   "PopUps_DB_1".Absolute_Encoder[#HMI_No].AE_Position_1 := "Control_DB".VTD_Sys[#Sys_No].Inputs.AE_Position_1;
   "PopUps_DB_1".Absolute_Encoder[#HMI_No].AE_Position_2 := "Control_DB".VTD_Sys[#Sys_No].Inputs.AE_Position_2;
   "PopUps_DB_1".Absolute_Encoder[#HMI_No].AE_Speed := "Control_DB".VTD_Sys[#Sys_No].Inputs.AE_Speed;
   "PopUps_DB_1".Absolute_Encoder[#HMI_No].AE_Status_1 := "Control_DB".VTD_Sys[#Sys_No].Inputs.AE_Status_1;
   "PopUps_DB_1".Absolute_Encoder[#HMI_No].AE_Status_2 := "Control_DB".VTD_Sys[#Sys_No].Inputs.AE_Status_2;

   //Instruction
   IF NOT "VTD_HMI".Charge_VTD_Commands[#HMI_No] THEN
       "Control_DB".VTD_Sys[#Sys_No].Instruction.Reset := "VTD_HMI".Reset[#HMI_No] OR "Screen_DB_1".Reset_All[#HMI_No];
       "Control_DB".VTD_Sys[#Sys_No].Instruction.Enable := "VTD_HMI".Enable[#HMI_No];
       IF "VTD_HMI".Stop[#HMI_No] THEN
           "Control_DB".VTD_Sys[#Sys_No].Instruction.Stop := TRUE;
       ELSIF "Screen_DB_1".Reset_All[1] OR "VTD_HMI".Reset[#HMI_No] THEN
           "Control_DB".VTD_Sys[#Sys_No].Instruction.Stop := "VTD_HMI".Stop[#HMI_No] := FALSE;
       END_IF;

       IF "Control_DB".VTD_Sys[#Sys_No].Mode <> 3 THEN
           "Control_DB".VTD_Sys[#Sys_No].Instruction.Pallet_Type := "VTD_HMI".Pallet_Type[#HMI_No];
           "Control_DB".VTD_Sys[#Sys_No].Instruction.Task_ID := "VTD_HMI".Task_ID[#HMI_No];

           IF "Control_DB".VTD_Sys[#Sys_No].Mode = 2 AND "VTD_HMI".Move_To_Level[#HMI_No] <> 0 THEN
               "Control_DB".VTD_Sys[#Sys_No].Instruction.Move_To_Level := "VTD_HMI".Move_To_Level[#HMI_No];
               "VTD_HMI".Move_To_Level[#HMI_No] := 0;
           END_IF;

           //UP
           IF "Control_DB".VTD_Sys[#Sys_No].LE < "Settings_DB".VTD_Sys[#Sys_No].Teach_Values.Levels_LE[#HMI_Box MOD 10 + 1] - 150
           THEN
               "Control_DB".VTD_Sys[#Sys_No].Instruction.Manual_Up := "VTD_HMI".Manual_Up[#HMI_No];
           ELSE
               "Control_DB".VTD_Sys[#Sys_No].Instruction.Manual_Up := "VTD_HMI".Manual_Up[#HMI_No] := FALSE;
           END_IF;
           //DOWN
           IF "Control_DB".VTD_Sys[#Sys_No].LE > "Settings_DB".VTD_Sys[#Sys_No].Teach_Values.Levels_LE[#HMI_Box MOD 10]
           THEN
               "Control_DB".VTD_Sys[#Sys_No].Instruction.Manual_Down := "VTD_HMI".Manual_Down[#HMI_No];
           ELSE
               "Control_DB".VTD_Sys[#Sys_No].Instruction.Manual_Down := "VTD_HMI".Manual_Down[#HMI_No] := FALSE;
           END_IF;

           "Control_DB".VTD_Sys[#Sys_No].Instruction.Manual_LP_Retract := "VTD_HMI".Manual_DP_Retract[#HMI_No];
           "Control_DB".VTD_Sys[#Sys_No].Instruction.Manual_LP_Extend := "VTD_HMI".Manual_DP_Extend[#HMI_No];
       END_IF;

       //ABSOLUTE ENCODER
       "Control_DB".VTD_Sys[#Sys_No].Outputs.AE_Control_Word_1 := "PopUps_DB_1".Absolute_Encoder[#HMI_No].AE_Control_Word_1;
       "Control_DB".VTD_Sys[#Sys_No].Outputs.AE_Control_Word_2 := "PopUps_DB_1".Absolute_Encoder[#HMI_No].AE_Control_Word_2;

       //LINEAR ENCODER
       "VTD_HMI".LE_Bypass[#Sys_No] := "PopUps_DB_1".Linear_Encoder[#HMI_No].LE_Bypass;

       //BARCODE
       #BCD_Start_Comm_Test_HMI := "PopUps_DB_1".Lector_Barcode[#HMI_No].BCD_Test_Comm;
       #BCD_Enable_Trigger_HMI  := "PopUps_DB_1".Lector_Barcode[#HMI_No].BCD_Enable_Trigger;
       #BCD_Disable_Trigger_HMI   := "PopUps_DB_1".Lector_Barcode[#HMI_No].BCD_Disable_Trigger;
       #BCD_Execute_Function  := "PopUps_DB_1".Lector_Barcode[#HMI_No].BCD_Execute_Function;
   END_IF;
END_FUNCTION

FUNCTION "FindBoolField" : Bool   // FC17, SCL
{ S7_Optimized_Access := 'TRUE' }
VERSION : 0.1
// stored: AutoNumber true, IsIECCheckEnabled false, SetENOAutomatically false, UDAEnableTagReadback false
   VAR_INPUT
      FieldName : String;
      JsonStr : String;
   END_VAR
   VAR_TEMP
      searchStr : String;
      foundPos : Int;
      valueStr : String;
      afterField : String;
      bResult : Bool;
   END_VAR
BEGIN
   // Build search string
   #searchStr := CONCAT(IN1 := '"', IN2 := #FieldName);
   #searchStr := CONCAT(IN1 := #searchStr, IN2 := '" :');

   // Serach for JSON field
   #foundPos := FIND(IN1 := #JsonStr, IN2 := #searchStr);

   IF #foundPos > 0 THEN
       // Take to 20 characters after the field
       #afterField := MID(IN := #JsonStr, P := #foundPos + LEN(#searchStr), L := 20);

       // Normalize to remove whitespace if necessary
       // (or compare directly)
       IF FIND(IN1 := #afterField, IN2 := 'true') > 0 THEN
           #bResult := TRUE;
       ELSIF FIND(IN1 := #afterField, IN2 := 'false') > 0 THEN
           #bResult := FALSE;
       ELSE
           #bResult := FALSE; // default if value not found
       END_IF;
   ELSE
       #bResult := FALSE;
   END_IF;

   #FindBoolField := #bResult;
END_FUNCTION

FUNCTION "FindDINTFieldFragmented" : DInt   // FC20, SCL
{ S7_Optimized_Access := 'TRUE' }
VERSION : 0.1
// stored: AutoNumber true, IsIECCheckEnabled false, SetENOAutomatically false, UDAEnableTagReadback false
   VAR_INPUT
      FieldName : String;
      Str1 : String;
      Str2 : String;
   END_VAR
   VAR_TEMP
      searchStr : String;
      iStart : Int;
      iEnd : Int;
      tempVal : String;
      fieldFound : Bool;
      loopIdx : Int;
   END_VAR
BEGIN
   // Build search string
   #searchStr := CONCAT(IN1 := '"', IN2 := #FieldName);
   #searchStr := CONCAT(IN1 := #searchStr, IN2 := '" :');

   // Serach for JSON field
   #iStart := FIND(IN1 := #Str1, IN2 := #searchStr);

   IF #iStart > 0 THEN
       // Found full field in String_1
       #iEnd := FIND(IN1 := MID(IN := #Str1, P := #iStart + LEN(#searchStr), L := 20), IN2 := ',');
       IF #iEnd = 0 THEN
           #iEnd := FIND(IN1 := MID(IN := #Str1, P := #iStart + LEN(#searchStr), L := 20), IN2 := '}');
       END_IF;
       IF #iEnd > 0 THEN
           #tempVal := MID(IN := #Str1, P := #iStart + LEN(#searchStr), L := #iEnd - 1);
           #fieldFound := TRUE;
       END_IF;
   END_IF;

   // Search for full field in Str2
   IF NOT #fieldFound THEN
       #iStart := FIND(IN1 := #Str2, IN2 := #searchStr);
       IF #iStart > 0 THEN
           #iEnd := FIND(IN1 := MID(IN := #Str2, P := #iStart + LEN(#searchStr), L := 20), IN2 := ',');
           IF #iEnd = 0 THEN
               #iEnd := FIND(IN1 := MID(IN := #Str2, P := #iStart + LEN(#searchStr), L := 20), IN2 := '}');
           END_IF;
           IF #iEnd > 0 THEN
               #tempVal := MID(IN := #Str2, P := #iStart + LEN(#searchStr), L := #iEnd - 1);
               #fieldFound := TRUE;
           END_IF;
       END_IF;
   END_IF;

   // Search for fragmented field: end of name in Str1 and beginning in Str2
   IF NOT #fieldFound THEN
       // Examines last 10 characters of String_1
       FOR #loopIdx := LEN(#Str1) - 15 TO LEN(#Str1) DO
           IF MID(IN := #Str1, P := #loopIdx, L := 1) = '"' THEN
               #tempVal := MID(IN := #Str1, P := #loopIdx, L := LEN(#Str1) - #loopIdx + 1);
               #tempVal := CONCAT(IN1 := #tempVal, IN2 := #Str2); // concatenates piece from beginning of String_2
               #iStart := FIND(IN1 := #tempVal, IN2 := #searchStr);
               IF #iStart > 0 THEN
                   #iEnd := FIND(IN1 := MID(IN := #tempVal, P := #iStart + LEN(#searchStr), L := 20), IN2 := ',');
                   IF #iEnd = 0 THEN
                       #iEnd := FIND(IN1 := MID(IN := #tempVal, P := #iStart + LEN(#searchStr), L := 20), IN2 := '}');
                   END_IF;
                   IF #iEnd > 0 THEN
                       #tempVal := MID(IN := #tempVal, P := #iStart + LEN(#searchStr), L := #iEnd - 1);
                       #fieldFound := TRUE;
                   END_IF;
               END_IF;
               EXIT; // found, you can leave
           END_IF;
       END_FOR;
   END_IF;

   // Return value
   IF #fieldFound THEN
       #FindDINTFieldFragmented := STRING_TO_DINT(#tempVal);
   ELSE
       #FindDINTFieldFragmented := -9999; // default value if not found
   END_IF;
END_FUNCTION

FUNCTION "FindINTFieldFragmented" : Int   // FC22, SCL
{ S7_Optimized_Access := 'TRUE' }
VERSION : 0.1
// stored: AutoNumber true, IsIECCheckEnabled false, SetENOAutomatically false, UDAEnableTagReadback false
   VAR_INPUT
      FieldName : String;
      Str1 : String;
      Str2 : String;
   END_VAR
   VAR_TEMP
      searchStr : String;
      iStart : Int;
      iEnd : Int;
      tempVal : String;
      fieldFound : Bool;
      loopIdx : Int;
   END_VAR
BEGIN
   // Build search string
   #searchStr := CONCAT(IN1 := '"', IN2 := #FieldName);
   #searchStr := CONCAT(IN1 := #searchStr, IN2 := '" :');

   // Serach for JSON field
   #iStart := FIND(IN1 := #Str1, IN2 := #searchStr);

   IF #iStart > 0 THEN
       // Found full field in String_1
       #iEnd := FIND(IN1 := MID(IN := #Str1, P := #iStart + LEN(#searchStr), L := 20), IN2 := ',');
       IF #iEnd = 0 THEN
           #iEnd := FIND(IN1 := MID(IN := #Str1, P := #iStart + LEN(#searchStr), L := 20), IN2 := '}');
       END_IF;
       IF #iEnd > 0 THEN
           #tempVal := MID(IN := #Str1, P := #iStart + LEN(#searchStr), L := #iEnd - 1);
           #fieldFound := TRUE;
       END_IF;
   END_IF;

   // Search for full field in Str2
   IF NOT #fieldFound THEN
       #iStart := FIND(IN1 := #Str2, IN2 := #searchStr);
       IF #iStart > 0 THEN
           #iEnd := FIND(IN1 := MID(IN := #Str2, P := #iStart + LEN(#searchStr), L := 20), IN2 := ',');
           IF #iEnd = 0 THEN
               #iEnd := FIND(IN1 := MID(IN := #Str2, P := #iStart + LEN(#searchStr), L := 20), IN2 := '}');
           END_IF;
           IF #iEnd > 0 THEN
               #tempVal := MID(IN := #Str2, P := #iStart + LEN(#searchStr), L := #iEnd - 1);
               #fieldFound := TRUE;
           END_IF;
       END_IF;
   END_IF;

   // Search for fragmented field: end of name in Str1 and beginning in Str2
   IF NOT #fieldFound THEN
       // Examines last 10 characters of String_1
       FOR #loopIdx := LEN(#Str1) - 15 TO LEN(#Str1) DO
           IF MID(IN := #Str1, P := #loopIdx, L := 1) = '"' THEN
               #tempVal := MID(IN := #Str1, P := #loopIdx, L := LEN(#Str1) - #loopIdx + 1);
               #tempVal := CONCAT(IN1 := #tempVal, IN2 := #Str2); // concatenates piece from beginning of String_2
               #iStart := FIND(IN1 := #tempVal, IN2 := #searchStr);
               IF #iStart > 0 THEN
                   #iEnd := FIND(IN1 := MID(IN := #tempVal, P := #iStart + LEN(#searchStr), L := 20), IN2 := ',');
                   IF #iEnd = 0 THEN
                       #iEnd := FIND(IN1 := MID(IN := #tempVal, P := #iStart + LEN(#searchStr), L := 20), IN2 := '}');
                   END_IF;
                   IF #iEnd > 0 THEN
                       #tempVal := MID(IN := #tempVal, P := #iStart + LEN(#searchStr), L := #iEnd - 1);
                       #fieldFound := TRUE;
                   END_IF;
               END_IF;
               EXIT; // found, you can leave
           END_IF;
       END_FOR;
   END_IF;

   // Return value
   IF #fieldFound THEN
       #FindINTFieldFragmented := STRING_TO_INT(#tempVal);
   ELSE
       #FindINTFieldFragmented := -9999; // default value if not found
   END_IF;
END_FUNCTION

FUNCTION "FindIntField" : Int   // FC18, SCL
{ S7_Optimized_Access := 'TRUE' }
VERSION : 0.1
// stored: AutoNumber true, IsIECCheckEnabled false, SetENOAutomatically false, UDAEnableTagReadback false
   VAR_INPUT
      FieldName : String;
      JsonStr : String;
   END_VAR
   VAR_TEMP
      searchStr : String;
      foundPos : Int;
      valueStr : String;
      delimPos : Int;
   END_VAR
BEGIN
   // Set up the search pattern, e.g. '"id":'
   #searchStr := CONCAT(IN1 := '"', IN2 := #FieldName);
   #searchStr := CONCAT(IN1 := #searchStr, IN2 := '" :');

   // Search the field
   #foundPos := FIND(IN1 := #JsonStr, IN2 := #searchStr);

   IF #foundPos > 0 THEN
       // Try to find a comma after the value
       #delimPos := FIND(
                         IN1 := MID(IN := #JsonStr, P := #foundPos + LEN(#searchStr), L := 10),
                         IN2 := ','
       );

       // If there is no comma, try to find the closing brace '}'
       IF #delimPos = 0 THEN
           #delimPos := FIND(
                             IN1 := MID(IN := #JsonStr, P := #foundPos + LEN(#searchStr), L := 10),
                             IN2 := '}'
           );
       END_IF;

       // If you find the end of value, extract the value
       IF #delimPos > 0 THEN
           #valueStr := MID(
                            IN := #JsonStr,
                            P := #foundPos + LEN(#searchStr),
                            L := #delimPos - 1
           );
           #FindIntField := STRING_TO_INT(#valueStr);
           RETURN;
       END_IF;
   END_IF;

   // Default return if not found or error
   #FindIntField := -9999;
END_FUNCTION

FUNCTION "FindSTRINGFieldFragmented" : String   // FC21, SCL
{ S7_Optimized_Access := 'TRUE' }
VERSION : 0.1
// stored: AutoNumber true, IsIECCheckEnabled false, SetENOAutomatically false, UDAEnableTagReadback false
   VAR_INPUT
      FieldName : String;
      Str1 : String;
      Str2 : String;
   END_VAR
   VAR_TEMP
      searchStr : String;
      iStart : Int;
      iEnd : Int;
      tempVal : String;
      fieldFound : Bool;
      loopIdx : Int;
   END_VAR
BEGIN
   // Build search string
   #searchStr := CONCAT(IN1 := '"', IN2 := #FieldName);
   #searchStr := CONCAT(IN1 := #searchStr, IN2 := '" :');

   // Serach for JSON field
   #iStart := FIND(IN1 := #Str1, IN2 := #searchStr);

   IF #iStart > 0 THEN
       // Found full field in String_1
       #iEnd := FIND(IN1 := MID(IN := #Str1, P := #iStart + LEN(#searchStr), L := 20), IN2 := ',');
       IF #iEnd = 0 THEN
           #iEnd := FIND(IN1 := MID(IN := #Str1, P := #iStart + LEN(#searchStr), L := 20), IN2 := '}');
       END_IF;
       IF #iEnd > 0 THEN
           #tempVal := MID(IN := #Str1, P := #iStart + LEN(#searchStr), L := #iEnd - 1);
           #fieldFound := TRUE;
       END_IF;
   END_IF;

   // Search for full field in Str2
   IF NOT #fieldFound THEN
       #iStart := FIND(IN1 := #Str2, IN2 := #searchStr);
       IF #iStart > 0 THEN
           #iEnd := FIND(IN1 := MID(IN := #Str2, P := #iStart + LEN(#searchStr), L := 20), IN2 := ',');
           IF #iEnd = 0 THEN
               #iEnd := FIND(IN1 := MID(IN := #Str2, P := #iStart + LEN(#searchStr), L := 20), IN2 := '}');
           END_IF;
           IF #iEnd > 0 THEN
               #tempVal := MID(IN := #Str2, P := #iStart + LEN(#searchStr), L := #iEnd - 1);
               #fieldFound := TRUE;
           END_IF;
       END_IF;
   END_IF;

   // Search for fragmented field: end of name in Str1 and beginning in Str2
   IF NOT #fieldFound THEN
       // Examines last 10 characters of String_1
       FOR #loopIdx := LEN(#Str1) - 15 TO LEN(#Str1) DO
           IF MID(IN := #Str1, P := #loopIdx, L := 1) = '"' THEN
               #tempVal := MID(IN := #Str1, P := #loopIdx, L := LEN(#Str1) - #loopIdx + 1);
               #tempVal := CONCAT(IN1 := #tempVal, IN2 := #Str2); // concatenates piece from beginning of String_2
               #iStart := FIND(IN1 := #tempVal, IN2 := #searchStr);
               IF #iStart > 0 THEN
                   #iEnd := FIND(IN1 := MID(IN := #tempVal, P := #iStart + LEN(#searchStr), L := 20), IN2 := ',');
                   IF #iEnd = 0 THEN
                       #iEnd := FIND(IN1 := MID(IN := #tempVal, P := #iStart + LEN(#searchStr), L := 20), IN2 := '}');
                   END_IF;
                   IF #iEnd > 0 THEN
                       #tempVal := MID(IN := #tempVal, P := #iStart + LEN(#searchStr), L := #iEnd - 1);
                       #fieldFound := TRUE;
                   END_IF;
               END_IF;
               EXIT; // found, you can leave
           END_IF;
       END_FOR;
   END_IF;

   // Return value
   IF #fieldFound THEN
       #FindSTRINGFieldFragmented := #tempVal;
   ELSE
       #FindSTRINGFieldFragmented := 'NOT FOUND'; // default value if not found
   END_IF;
END_FUNCTION

FUNCTION "FindStringField" : String   // FC19, SCL
{ S7_Optimized_Access := 'TRUE' }
VERSION : 0.1
// stored: AutoNumber true, IsIECCheckEnabled false, SetENOAutomatically false, UDAEnableTagReadback false
   VAR_INPUT
      FieldName : String;
      JsonStr : String;
   END_VAR
   VAR_TEMP
      searchStr : String;
      foundPos : Int;
      resultStr : String;
      quotePos1 : Int;
      quotePos2 : Int;
   END_VAR
BEGIN
   // Sets search pattern → ex: '"loadstate":'
   #searchStr := CONCAT(IN1 := '"', IN2 := #FieldName);
   #searchStr := CONCAT(IN1 := #searchStr, IN2 := '" :');

   // Search in JSON
   #foundPos := FIND(IN1 := #JsonStr, IN2 := #searchStr);

   IF #foundPos > 0 THEN
       // Finds first quote after field
       #quotePos1 := FIND(IN1 := MID(IN := #JsonStr, P := #foundPos + LEN(#searchStr), L := 20), IN2 := '"');

       IF #quotePos1 > 0 THEN
           // Finds second quote after the first
           #quotePos2 := FIND(
                              IN1 := MID(IN := #JsonStr, P := #foundPos + LEN(IN := #searchStr) + #quotePos1, L := 10),
                              IN2 := '"'
           );

           IF #quotePos2 > 0 THEN
               #resultStr := MID(
                                 IN := #JsonStr,
                                 P := #foundPos + LEN(#searchStr) + #quotePos1,
                                 L := #quotePos2 - 1
               );
               #FindStringField := #resultStr;
               RETURN;
           END_IF;
       END_IF;
   END_IF;

   // If not found, returns empty string
   #FindStringField := '';
END_FUNCTION

FUNCTION "Gate_Status_Update_FC" : Void   // FC49, SCL
{ S7_Optimized_Access := 'TRUE' }
VERSION : 0.1
// stored: AutoNumber true, IsIECCheckEnabled false, SetENOAutomatically false, UDAEnableTagReadback false
   VAR_INPUT
      Gate_Index : Int;
      Request_Access : Bool;
      Stop_Mode_Granted : Bool;
   END_VAR
   VAR_OUTPUT
      DB_SM_To_LGX_Gate_Status : Array[0..10] of Byte;
   END_VAR
   VAR_TEMP
      tGateByte : Byte;
   END_VAR
BEGIN
   #tGateByte := 0;

   IF #Request_Access THEN
       #tGateByte := #tGateByte OR BYTE#16#01;
   END_IF; // Bit 0
   IF #Stop_Mode_Granted THEN
       #tGateByte := #tGateByte OR BYTE#16#02;
   END_IF; // Bit 1
   // Bits 2..7: Free

   IF #Gate_Index >= 0 AND #Gate_Index <= 10 THEN
       #DB_SM_To_LGX_Gate_Status[#Gate_Index] := #tGateByte;
   END_IF;
END_FUNCTION

FUNCTION "HMI_SAFETY_FC" : Void   // FC43, F_FBD
{ S7_Optimized_Access := 'TRUE' }
VERSION : 0.1
// stored: AutoNumber true, IsIECCheckEnabled false, UDAEnableTagReadback false
   VAR_INPUT
      HMI_Box_Connected : Int;
      HMI_Reset : Bool;
      HMI_EStop : Bool;
      HMI_Profinet_Error : Bool;
      Local_Mode : Bool;
   END_VAR
   VAR_OUTPUT
      HMI_Estop_Pressed_1 : Bool;
      HMI_Estop_Pressed_2 : Bool;
      HMI_Estop_Pressed_3 : Bool;
      HMI_Estop_Pressed_4 : Bool;
      HMI_Estop_Pressed_5 : Bool;
      Reset_Comissioning_1 : Bool;
      Reset_Comissioning_2 : Bool;
      Reset_Comissioning_3 : Bool;
      Reset_Comissioning_4 : Bool;
      Reset_Comissioning_5 : Bool;
   END_VAR
   VAR_TEMP   // added for the SCL form of the ladder/FBD networks
      _w1 : Bool;
   END_VAR
BEGIN

REGION Network 1: HMI CONNECTED IN THE SYSTEM 1
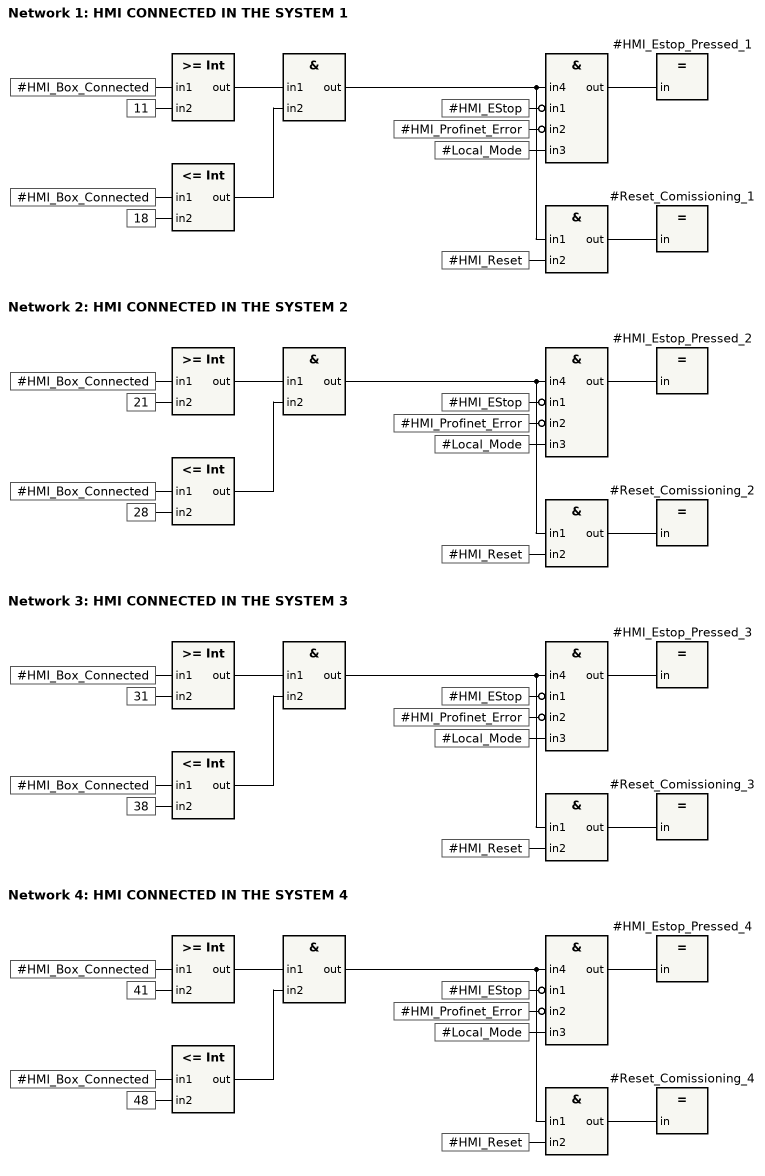
   #_w1 := (#HMI_Box_Connected >= 11) AND (#HMI_Box_Connected <= 18);
   #HMI_Estop_Pressed_1 := #_w1 AND NOT #HMI_EStop AND NOT #HMI_Profinet_Error AND #Local_Mode;
   #Reset_Comissioning_1 := #_w1 AND #HMI_Reset;
END_REGION

REGION Network 2: HMI CONNECTED IN THE SYSTEM 2
   #_w1 := (#HMI_Box_Connected >= 21) AND (#HMI_Box_Connected <= 28);
   #HMI_Estop_Pressed_2 := #_w1 AND NOT #HMI_EStop AND NOT #HMI_Profinet_Error AND #Local_Mode;
   #Reset_Comissioning_2 := #_w1 AND #HMI_Reset;
END_REGION

REGION Network 3: HMI CONNECTED IN THE SYSTEM 3
   #_w1 := (#HMI_Box_Connected >= 31) AND (#HMI_Box_Connected <= 38);
   #HMI_Estop_Pressed_3 := #_w1 AND NOT #HMI_EStop AND NOT #HMI_Profinet_Error AND #Local_Mode;
   #Reset_Comissioning_3 := #_w1 AND #HMI_Reset;
END_REGION

REGION Network 4: HMI CONNECTED IN THE SYSTEM 4
   #_w1 := (#HMI_Box_Connected >= 41) AND (#HMI_Box_Connected <= 48);
   #HMI_Estop_Pressed_4 := #_w1 AND NOT #HMI_EStop AND NOT #HMI_Profinet_Error AND #Local_Mode;
   #Reset_Comissioning_4 := #_w1 AND #HMI_Reset;
END_REGION

REGION Network 5: HMI CONNECTED IN THE SYSTEM 5
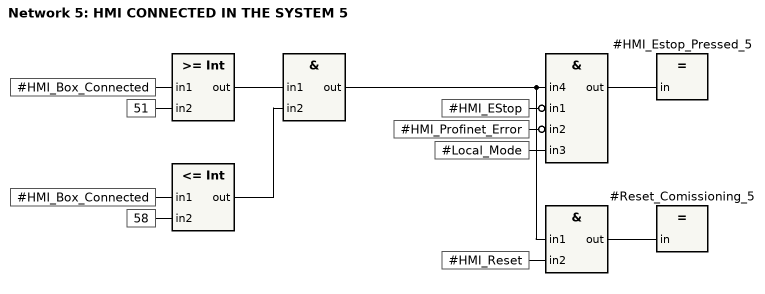
   #_w1 := (#HMI_Box_Connected >= 51) AND (#HMI_Box_Connected <= 58);
   #HMI_Estop_Pressed_5 := #_w1 AND NOT #HMI_EStop AND NOT #HMI_Profinet_Error AND #Local_Mode;
   #Reset_Comissioning_5 := #_w1 AND #HMI_Reset;
END_REGION
END_FUNCTION

FUNCTION "Handshake_Infeed_FC" : Void   // FC47, SCL
{ S7_Optimized_Access := 'TRUE' }
VERSION : 0.1
// stored: AutoNumber true, IsIECCheckEnabled false, SetENOAutomatically false, UDAEnableTagReadback false
   VAR_INPUT
      Infeed_Stop_Sensor : Bool;
      Ready_To_Receive : Bool;
      Auto_Mode : Bool;
      Transfer_In_Progress : Bool;
      DB_LGX_To_SM_Infeed_Ready_To_Send : Bool;
      DB_LGX_To_SM_Infeed_Transfer_In_Progress : Bool;
   END_VAR
   VAR_OUTPUT
      Fault_Handshake : Bool;
      DB_SM_To_LGX_Infeed_Ready_To_Receive : Bool;
      DB_SM_To_LGX_Infeed_Pallet_Received : Bool;
      DB_SM_To_LGX_Infeed_Transfer_In_Progress : Bool;
   END_VAR
   VAR_TEMP
      tReady_To_Receive_Condition : Bool;
      tPallet_Received_Condition : Bool;
   END_VAR
BEGIN
   // ---------------------------------------------------------
   // STEP 1: Is SM ready to receive?
   // Condition: SM in Auto, infeed conveyor healthy,
   //            no transfer in progress, no alarm
   // ---------------------------------------------------------
   #tReady_To_Receive_Condition :=
   #Auto_Mode
   AND #Ready_To_Receive
   AND NOT #DB_SM_To_LGX_Infeed_Ready_To_Receive
   AND NOT #DB_SM_To_LGX_Infeed_Pallet_Received;

   IF #DB_LGX_To_SM_Infeed_Ready_To_Send
       AND #tReady_To_Receive_Condition THEN
       #DB_SM_To_LGX_Infeed_Ready_To_Receive := TRUE;
   END_IF;

   // ---------------------------------------------------------
   // STEP 2: Confirm pallet received
   // Condition: Photocell active while transfer is in progress
   // ---------------------------------------------------------
   // #tPallet_Received_Condition :=
   // #Infeed_Stop_Sensor
   // AND #DB_LGX_To_SM_Infeed_Transfer_In_Progress
   // AND #DB_SM_To_LGX_Infeed_Ready_To_Receive;
   // 
   #tPallet_Received_Condition :=
   #Infeed_Stop_Sensor;

   IF #tPallet_Received_Condition THEN
       #DB_SM_To_LGX_Infeed_Pallet_Received := TRUE;
       #DB_SM_To_LGX_Infeed_Ready_To_Receive := FALSE;
   ELSE
       #DB_SM_To_LGX_Infeed_Pallet_Received := FALSE;
   END_IF;

   // ---------------------------------------------------------
   // STEP 3: Reset after LGX confirms end of transfer
   // (LGX resets Transfer_In_Progress upon receiving Pallet_Received)
   // ---------------------------------------------------------
   // IF #DB_SM_To_LGX_Infeed_Pallet_Received
   //     AND NOT #DB_LGX_To_SM_Infeed_Transfer_In_Progress THEN
   //     #DB_SM_To_LGX_Infeed_Pallet_Received := FALSE;
   // END_IF;

   // ---------------------------------------------------------
   // STEP 4: Reset Ready_To_Receive if LGX withdraws Ready_To_Send
   // (e.g. LGX cancelled the operation before starting transfer)
   // ---------------------------------------------------------
   IF NOT #DB_LGX_To_SM_Infeed_Ready_To_Send
       AND NOT #DB_LGX_To_SM_Infeed_Transfer_In_Progress THEN
       #DB_SM_To_LGX_Infeed_Ready_To_Receive := FALSE;
   END_IF;

   // ---------------------------------------------------------
   // FAULT SUPERVISION
   // If Transfer_In_Progress remains active without pallet arriving:
   // use external timer / timeout bit (implement in OB1)
   // ---------------------------------------------------------
   #Fault_Handshake := FALSE; // Placeholder - implement watchdog

   #DB_SM_To_LGX_Infeed_Transfer_In_Progress := #Transfer_In_Progress;
END_FUNCTION

FUNCTION "Handshake_Outfeed_FC" : Void   // FC51, SCL
{ S7_Optimized_Access := 'TRUE' }
VERSION : 0.1
// stored: AutoNumber true, IsIECCheckEnabled false, SetENOAutomatically false, UDAEnableTagReadback false
   VAR_INPUT
      Auto_Mode : Bool;
      Ready_To_Send : Bool;
      Conv_Occupied : Bool;
      Transfer_In_Progress : Bool;
      DB_LGX_To_SM_Outfeed_Ready_To_Receive : Bool;
   END_VAR
   VAR_OUTPUT
      Fault_Handshake : Bool;
      DB_SM_To_LGX_Outfeed_Transfer_In_Progress : Bool;
      DB_SM_To_LGX_Outfeed_Ocuppied : Bool;
      DB_SM_To_LGX_Outfeed_Ready_To_Send : Bool;
   END_VAR
   VAR_TEMP
      tCanSend : Bool;
   END_VAR
BEGIN
   // ---------------------------------------------------------
   // STEP 1: Is SM ready to send?
   // Condition: pallet waiting at exit, SM in auto,
   //            no transfer in progress
   // ---------------------------------------------------------
   #tCanSend :=
   #Auto_Mode
   AND #Conv_Occupied
   AND #Ready_To_Send
   AND NOT #DB_SM_To_LGX_Outfeed_Transfer_In_Progress;

   IF #tCanSend
       AND NOT #DB_SM_To_LGX_Outfeed_Ready_To_Send THEN
       #DB_SM_To_LGX_Outfeed_Ready_To_Send := TRUE;
   END_IF;

   // ---------------------------------------------------------
   // STEP 2: LGX responded Ready_To_Receive → start transfer
   // ---------------------------------------------------------
   IF NOT #Conv_Occupied THEN
       // #DB_SM_To_LGX_Outfeed_Transfer_In_Progress := TRUE;
       #DB_SM_To_LGX_Outfeed_Ready_To_Send := FALSE;
   END_IF;

   // ---------------------------------------------------------
   // STEP 3: LGX confirmed pallet received
   // → SM resets Transfer_In_Progress
   // ---------------------------------------------------------
   // IF #DB_SM_To_LGX_Outfeed_Transfer_In_Progress
   //     AND #DB_LGX_To_SM_Outfeed_Ready_To_Receive THEN
   //     #DB_SM_To_LGX_Outfeed_Transfer_In_Progress := FALSE;
   // END_IF;

   #DB_SM_To_LGX_Outfeed_Transfer_In_Progress := #Transfer_In_Progress;
   #DB_SM_To_LGX_Outfeed_Ocuppied := #Conv_Occupied;
   // ---------------------------------------------------------
   // STEP 4: Reset Ready_To_Send if pallet removed or SM left auto mode
   // ---------------------------------------------------------
   IF NOT #Ready_To_Send OR NOT #Auto_Mode THEN
       IF NOT #DB_SM_To_LGX_Outfeed_Transfer_In_Progress THEN
           #DB_SM_To_LGX_Outfeed_Ready_To_Send := FALSE;
       END_IF;
   END_IF;

   #Fault_Handshake := FALSE; // Placeholder
END_FUNCTION

FUNCTION "ID_Decode_F" : Void   // FC3, SCL
{ S7_Optimized_Access := 'TRUE' }
VERSION : 0.1
// stored: AutoNumber true, IsIECCheckEnabled false, SetENOAutomatically false, UDAEnableTagReadback false
   VAR_INPUT
      ID : DInt;
   END_VAR
   VAR_IN_OUT
      ID_Decoded : "ID_Decoded";
   END_VAR
   VAR_TEMP
      Temp : UInt;
   END_VAR
BEGIN

   // Extract XX (first two digits)
   #ID_Decoded.Device_Type := #ID / 10000;        // 123456 / 10000 = 12

   // Extract YY (middle two digits)
   #ID_Decoded.Level := (#ID MOD 10000) / 100; // 123456 % 10000 = 3456 → 3456 / 100 = 34

   // Extract ZZ (last two digits)
   #ID_Decoded.VTD := #ID MOD 100;       // 123456 % 100 = 56
END_FUNCTION

FUNCTION "IsIPAddress" : Bool   // FC4, SCL
TITLE = IsIPAddress
{ S7_Optimized_Access := 'TRUE' }
VERSION : 0.1
// Evaluates whether a given String contains a valid IP address
// stored: AutoNumber true, IsIECCheckEnabled true, SetENOAutomatically true, UDAEnableTagReadback false
   VAR_INPUT
      address : String;   // Address to be evaluated
   END_VAR
   VAR_OUTPUT
      ipAddress : IP_V4;   // Parsed IP address if passed address is IP address
   END_VAR
   VAR_TEMP
      tempAddress : String;   // Passed address
      tempOctet : String;   // Current octet
      tempIndex : DInt;   // Index for loop
      tempPos : Int;   // Position of found separator
      tempNum : Int;   // Converted octet
      tempIp : IP_V4;   // Parsed IP address
   END_VAR
   VAR CONSTANT
      MAX_VALUE : USInt := 255;   // Max. valid value of octet
      NUM_OCTETS : DInt := 4;   // Number of octets
      CHAR_ZERO : Char := '0';   // ASCII character '0'
   END_VAR
   // Ret_Val : Return value
BEGIN
   REGION BLOCK INFO HEADER
     //===============================================================================
     // SIEMENS / (c)Copyright 2024
     //-------------------------------------------------------------------------------
     // Title:        IsIPAddress
     // Function:     Evaluates whether a given String contains a valid IP address
     // Library:      --
     // Author:       Siemens Industry Online Support
     // Tested with:  CPU 1515-2 PN V3.1
     // Engineering:  TIA Portal V17
     // Restrictions: --
     // Requirements: S7-1200 with firmware V4.4 or higher
     //               S7-1500 with firmware V2.0 or higher
     //-------------------------------------------------------------------------------
     // Change log table:
     // Version  | Date       | Expert in charge       | Changes applied
     //-------------------------------------------------------------------------------
     // 01.00.00 | 2024-02-12 | Online Support         | First released version
     //===============================================================================
   END_REGION

   #tempAddress := #address;
   #IsIPAddress := FALSE; // Will be overwritten if IP address is detected
   #ipAddress := #tempIp; // Zero output parameter

   FOR #tempIndex := 1 TO #NUM_OCTETS DO
     #tempPos := FIND(IN1 := #tempAddress, IN2 := '.'); // Find separator

     IF (#tempPos > 0 OR #tempIndex = #NUM_OCTETS) // Separator found with exception of last octet
       AND NOT (#tempPos > 0 AND #tempIndex = #NUM_OCTETS) // No separator found in last octet
       AND #tempPos <= 4 // 3  characters or less
     THEN
       IF #tempIndex < #NUM_OCTETS THEN // First three octets
         #tempOctet := LEFT(IN := #tempAddress, L := #tempPos - 1);
       ELSE// Last octet
         #tempOctet := #tempAddress;
       END_IF;

       STRG_VAL(IN := #tempOctet,
                FORMAT := 0,
                P := 1,
                OUT => #tempNum);

       IF #tempNum >= 0 AND #tempNum <= #MAX_VALUE // Within 0 and 255
         AND NOT (#tempNum = 0 AND #tempIndex = 1) // Not 0 in first octet
         AND NOT (#tempNum = 0 AND #tempOctet[1] <> #CHAR_ZERO) // Not 0 because of invalid character
       THEN
         #tempIp.ADDR[#tempIndex] := INT_TO_BYTE(#tempNum);
         #tempAddress := RIGHT(IN := #tempAddress, L := LEN(#tempAddress) - #tempPos); // Remove evaluated octet
       ELSE // Address is not IP address
         EXIT;
       END_IF;
     ELSE // Address is not IP address
       EXIT;
     END_IF;

     IF #tempIndex = #NUM_OCTETS THEN // End of loop reached, address is IP address
       #ipAddress := #tempIp;
       #IsIPAddress := true;
     END_IF;
   END_FOR;
END_FUNCTION

FUNCTION "LMQTT_ConvertToUtf8" : Void   // FC6, SCL
TITLE = LMQTT_ConvertToUtf8
{ S7_Optimized_Access := 'TRUE' }
AUTHOR : SIEMENS
FAMILY : LMQTT
VERSION : 1.0
// Function to convert a WCHAR to a UTF-8 conformant byte sequence
// stored: AutoNumber true, IsIECCheckEnabled true, SetENOAutomatically false, UDAEnableTagReadback false
   VAR_INPUT
      character : WChar;   // Character that shall be converted to UTF-8
   END_VAR
   VAR_OUTPUT
      convertedUtf8 : DWord;   // UTF-8 conformant byte sequence. B0 stores first Byte, B1 second and B2 third Byte. B3 is not used
      bytesUsed : USInt;   // Amount of Bytes converted. Ranges from 1 to 3.
      error : Bool;   // TRUE: An error occurred during the execution of the FC
      status : Word;   // 16#0000 - 16#7FFF: Status of the FC, 16#8000 - 16#FFFF: Error identification
   END_VAR
   VAR_TEMP
      tempStatus : Word;   // temp value for output 'status'
      tempConvertedUtf8 : DWord;   // temp value for output 'convertedUtf8'
      tempBytesUsed : USInt;   // temp value for output 'bytesUsed'
      tempCharacter : WChar;   // temp value for input 'character'
   END_VAR
   VAR CONSTANT
      STATUS_NO_ERROR : Word := 16#0000;   // no error status
      STATUS_EXECUTION_FINISHED : Word := 16#0000;   // Execution finished without errors
      ERR_UNDEFINED : Word := 16#8000;   // Error due to an undefined case
      USINT_NULL : USInt := 0;   // Init value with 0
      DWORD_NULL : DWord := 16#0000_0000;   // Init value with 0
      EMPTY_WCHAR : WChar := WCHAR#' ';   // Empty WChar for comparison
      BELOW_7F : Word := 16#007F;   // Upper limit for character if only one Byte used
      BELOW_7FF : Word := 16#07FF;   // Upper limit for character if two Byte used
      BELOW_MAX_FFFF : Word := 16#FFFF;   // Upper limit for character if three Byte used
      BYTE_3F : Byte := 16#3F;   // Conversion Value
      BYTE_80 : Byte := 16#80;   // Conversion Value
      BYTE_C0 : Byte := 16#C0;   // Conversion Value
      BYTE_E0 : Byte := 16#E0;   // Conversion Value
      USINT_ONE : USInt := 1;   // Const Value to assign amount of bytes used
      USINT_TWO : USInt := 2;   // Const Value to assign amount of bytes used
      USINT_THREE : USInt := 3;   // Const Value to assign amount of bytes used
   END_VAR
   // Ret_Val : No return for this FC - see error and status output
BEGIN
   REGION BLOCK INFO HEADER
       //=============================================================================
       // SIEMENS AG
       // (c)Copyright 2020
       //-----------------------------------------------------------------------------
       // Library:       LMQTT
       // Tested with:   CPU 1516-3 PN/DP V2.8
       // Engineering:   TIA Portal V16
       // Restrictions:  --
       // Requirements:  --
       // Functionality: Converts a single WChar Character to a valid UTF-8 encoded byte sequence and saves this to a DWord.
       //                The amount of bytes saved is stored in bytesUsed Output.
       //-----------------------------------------------------------------------------
       // Change log table:
       // Version    Date         Expert in charge         Changes applied
       // 03.00.00   01.10.2020   Siemens Online Support   First released version
       //=============================================================================
   END_REGION

   REGION INITIALISATION  
       // Initialize functionality: reset of variables, diagnostics, etc.
       #tempConvertedUtf8 := #DWORD_NULL;
       #tempBytesUsed := #USINT_NULL;
       #tempStatus := #STATUS_NO_ERROR;
       //assign temp value from input:
        #tempCharacter := #character;

   END_REGION

   REGION PROGRAM LOGIC
       // Use this region for application specific code
       IF #tempCharacter = #EMPTY_WCHAR THEN
           //will be only 1 byte occupied
           #tempConvertedUtf8 := WCHAR_TO_DWORD(#tempCharacter);
           #tempBytesUsed := #USINT_ONE;
       ELSIF (WCHAR_TO_WORD(#tempCharacter) <= (#BELOW_7F)) THEN
           //will be only 1 byte occupied
           #tempConvertedUtf8 := WCHAR_TO_DWORD(#tempCharacter);
           #tempBytesUsed := #USINT_ONE;
       ELSIF (WCHAR_TO_WORD(#tempCharacter) <= (#BELOW_7FF)) THEN
           //will be 2 byte occupied
           #tempConvertedUtf8.%B1 := (WCHAR_TO_BYTE(#tempCharacter) AND #BYTE_3F) OR #BYTE_80;
           #tempConvertedUtf8.%B0 := WORD_TO_BYTE(SHR(IN := WCHAR_TO_WORD(#tempCharacter), N := 6)) OR #BYTE_C0;
           #tempBytesUsed := #USINT_TWO;
       ELSIF (WCHAR_TO_WORD(#tempCharacter) <= (#BELOW_MAX_FFFF)) THEN
           //will be 3 byte occupied
           #tempConvertedUtf8.%B2 := (WCHAR_TO_BYTE(#tempCharacter) AND #BYTE_3F) OR #BYTE_80;
           #tempConvertedUtf8.%B1 := (WORD_TO_BYTE(SHR(IN := WCHAR_TO_WORD(#tempCharacter), N := 6)) AND #BYTE_3F) OR #BYTE_80;
           #tempConvertedUtf8.%B0 := WORD_TO_BYTE(SHR(IN := WCHAR_TO_WORD(#tempCharacter), N := 12)) OR #BYTE_E0;
           #tempBytesUsed := #USINT_THREE;
       END_IF;
   END_REGION

   REGION OUTPUTS
       // Write application specific temp values to outputs
       #bytesUsed := #tempBytesUsed;
       #convertedUtf8 := #tempConvertedUtf8;
       // Write error and status
       #error := #tempStatus.%X15;
       #status := #tempStatus;
       // ENO mechanism is not used --> ENO := TRUE;
       ENO := TRUE;
   END_REGION
END_FUNCTION

FUNCTION_BLOCK "Main_Panel"   // FB16, F_LAD
{ S7_Optimized_Access := 'TRUE' }
VERSION : 0.1
// stored: AutoNumber true, IsIECCheckEnabled false, UDAEnableTagReadback false
   VAR_INPUT
      Estop_Cabinet_Ch1 : Bool;
      Reset_Cabinet : Bool;
      Bypass : "F_Bypass_MainPanel";
   END_VAR
   VAR_OUTPUT
      Safety_OK : Bool;
      Main_Panel_OK : Bool;
      Bypass_Warning : Bool;
      ACK { ExternalAccessible := 'False'; ExternalVisible := 'False'; ExternalWritable := 'False'} : Bool;
   END_VAR
   VAR
      Estop_Cabinet_DB : ESTOP1;
   END_VAR
BEGIN

REGION Network 1: RESET CABINET
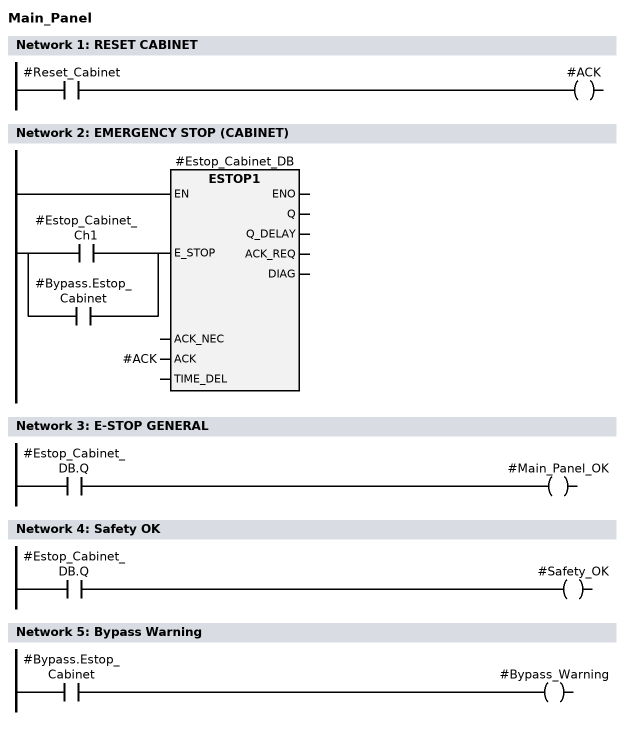
   RUNG wire#powerrail
      Contact( #Reset_Cabinet )
      Coil( #ACK )
   END_RUNG
   // the same network as SCL:
   #ACK := #Reset_Cabinet;
END_REGION

REGION Network 2: EMERGENCY STOP (CABINET)
   RUNG wire#powerrail
      #Estop_Cabinet_DB.ESTOP1(E_STOP := wire#w1, ACK_NEC :=, ACK := #ACK, TIME_DEL :=, Q =>, Q_DELAY =>, ACK_REQ =>, DIAG =>)
   END_RUNG
   RUNG wire#powerrail
      Contact( #Estop_Cabinet_Ch1 )
   END_RUNG wire#w1
   RUNG wire#powerrail
      Contact( #Bypass.Estop_Cabinet )
   END_RUNG wire#w1
   // the same network as SCL:
   #Estop_Cabinet_DB(E_STOP := #Estop_Cabinet_Ch1 OR #Bypass.Estop_Cabinet, ACK := #ACK);   // ESTOP1
END_REGION

REGION Network 3: E-STOP GENERAL
   RUNG wire#powerrail
      Contact( #Estop_Cabinet_DB.Q )
      Coil( #Main_Panel_OK )
   END_RUNG
   // the same network as SCL:
   #Main_Panel_OK := #Estop_Cabinet_DB.Q;
END_REGION

REGION Network 4: Safety OK
   RUNG wire#powerrail
      Contact( #Estop_Cabinet_DB.Q )
      Coil( #Safety_OK )
   END_RUNG
   // the same network as SCL:
   #Safety_OK := #Estop_Cabinet_DB.Q;
END_REGION

REGION Network 5: Bypass Warning
   RUNG wire#powerrail
      Contact( #Bypass.Estop_Cabinet )
      Coil( #Bypass_Warning )
   END_RUNG
   // the same network as SCL:
   #Bypass_Warning := #Bypass.Estop_Cabinet;
END_REGION
END_FUNCTION_BLOCK

FUNCTION_BLOCK "Main_Safety_RTG1"   // FB123, F_FBD
{ S7_Optimized_Access := 'TRUE' }
VERSION : 0.1
// stored: AutoNumber false, IsIECCheckEnabled false, UDAEnableTagReadback false
   VAR
      Safety_OK : Bool;
      ACK : Bool;
   END_VAR
   VAR_TEMP
      HMI_1_Estop_Pressed_1 : Bool;
      HMI_1_Estop_Pressed_2 : Bool;
      HMI_1_Estop_Pressed_3 : Bool;
      HMI_1_Estop_Pressed_4 : Bool;
      HMI_1_Estop_Pressed_5 : Bool;
      HMI_2_Estop_Pressed_1 : Bool;
      HMI_2_Estop_Pressed_2 : Bool;
      HMI_2_Estop_Pressed_3 : Bool;
      HMI_2_Estop_Pressed_4 : Bool;
      HMI_2_Estop_Pressed_5 : Bool;
      HMI_1_Reset_Comiss_1 : Bool;
      HMI_1_Reset_Comiss_2 : Bool;
      HMI_1_Reset_Comiss_3 : Bool;
      HMI_1_Reset_Comiss_4 : Bool;
      HMI_1_Reset_Comiss_5 : Bool;
      HMI_2_Reset_Comiss_1 : Bool;
      HMI_2_Reset_Comiss_2 : Bool;
      HMI_2_Reset_Comiss_3 : Bool;
      HMI_2_Reset_Comiss_4 : Bool;
      HMI_2_Reset_Comiss_5 : Bool;
   END_VAR
BEGIN

REGION Network 1: MAIN PANEL
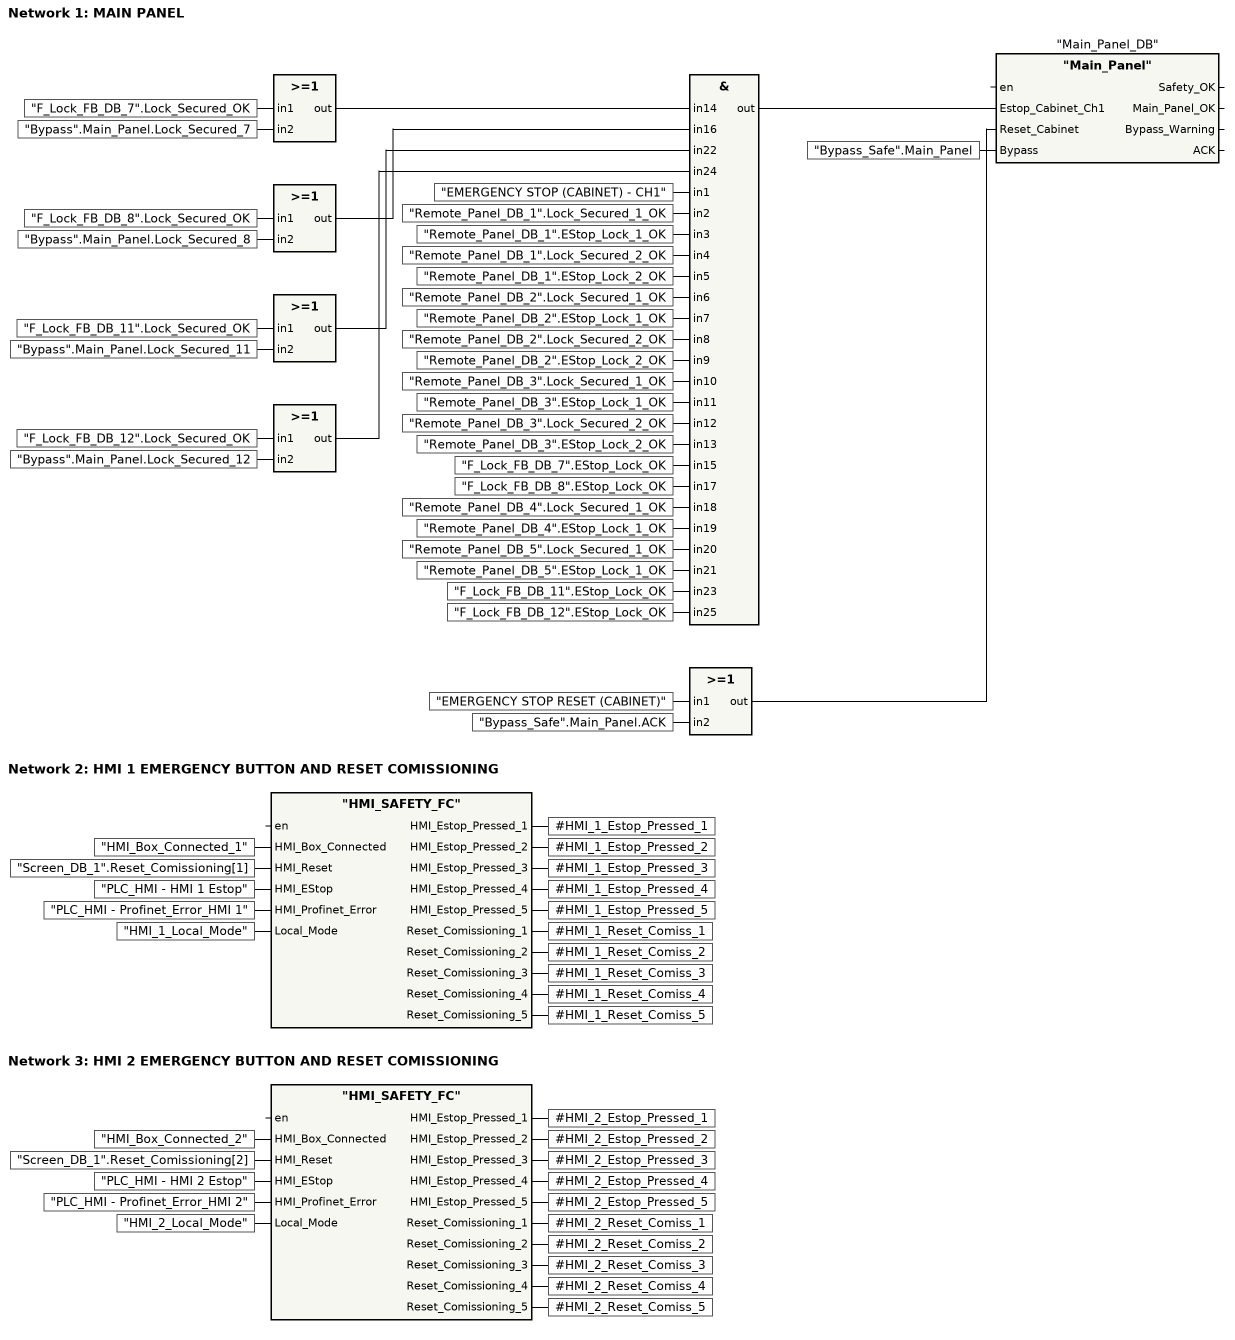
   "Main_Panel_DB"(Estop_Cabinet_Ch1 := ("F_Lock_FB_DB_7".Lock_Secured_OK OR "Bypass".Main_Panel.Lock_Secured_7) AND ("F_Lock_FB_DB_8".Lock_Secured_OK OR "Bypass".Main_Panel.Lock_Secured_8) AND ("F_Lock_FB_DB_11".Lock_Secured_OK OR "Bypass".Main_Panel.Lock_Secured_11) AND ("F_Lock_FB_DB_12".Lock_Secured_OK OR "Bypass".Main_Panel.Lock_Secured_12) AND "EMERGENCY STOP (CABINET) - CH1" AND "Remote_Panel_DB_1".Lock_Secured_1_OK AND "Remote_Panel_DB_1".EStop_Lock_1_OK AND "Remote_Panel_DB_1".Lock_Secured_2_OK AND "Remote_Panel_DB_1".EStop_Lock_2_OK AND "Remote_Panel_DB_2".Lock_Secured_1_OK AND "Remote_Panel_DB_2".EStop_Lock_1_OK AND "Remote_Panel_DB_2".Lock_Secured_2_OK AND "Remote_Panel_DB_2".EStop_Lock_2_OK AND "Remote_Panel_DB_3".Lock_Secured_1_OK AND "Remote_Panel_DB_3".EStop_Lock_1_OK AND "Remote_Panel_DB_3".Lock_Secured_2_OK AND "Remote_Panel_DB_3".EStop_Lock_2_OK AND "F_Lock_FB_DB_7".EStop_Lock_OK AND "F_Lock_FB_DB_8".EStop_Lock_OK AND "Remote_Panel_DB_4".Lock_Secured_1_OK AND "Remote_Panel_DB_4".EStop_Lock_1_OK AND "Remote_Panel_DB_5".Lock_Secured_1_OK AND "Remote_Panel_DB_5".EStop_Lock_1_OK AND "F_Lock_FB_DB_11".EStop_Lock_OK AND "F_Lock_FB_DB_12".EStop_Lock_OK,   // "Main_Panel"
                   Reset_Cabinet := "EMERGENCY STOP RESET (CABINET)" OR "Bypass_Safe".Main_Panel.ACK,
                   Bypass := "Bypass_Safe".Main_Panel);
END_REGION

REGION Network 2: HMI 1 EMERGENCY BUTTON AND RESET COMISSIONING
   "HMI_SAFETY_FC"(HMI_Box_Connected := "HMI_Box_Connected_1",
                   HMI_Reset := "Screen_DB_1".Reset_Comissioning[1],
                   HMI_EStop := "PLC_HMI - HMI 1 Estop",
                   HMI_Profinet_Error := "PLC_HMI - Profinet_Error_HMI 1",
                   Local_Mode := "HMI_1_Local_Mode",
                   HMI_Estop_Pressed_1 => #HMI_1_Estop_Pressed_1,
                   HMI_Estop_Pressed_2 => #HMI_1_Estop_Pressed_2,
                   HMI_Estop_Pressed_3 => #HMI_1_Estop_Pressed_3,
                   HMI_Estop_Pressed_4 => #HMI_1_Estop_Pressed_4,
                   HMI_Estop_Pressed_5 => #HMI_1_Estop_Pressed_5,
                   Reset_Comissioning_1 => #HMI_1_Reset_Comiss_1,
                   Reset_Comissioning_2 => #HMI_1_Reset_Comiss_2,
                   Reset_Comissioning_3 => #HMI_1_Reset_Comiss_3,
                   Reset_Comissioning_4 => #HMI_1_Reset_Comiss_4,
                   Reset_Comissioning_5 => #HMI_1_Reset_Comiss_5);
END_REGION

REGION Network 3: HMI 2 EMERGENCY BUTTON AND RESET COMISSIONING
   "HMI_SAFETY_FC"(HMI_Box_Connected := "HMI_Box_Connected_2",
                   HMI_Reset := "Screen_DB_1".Reset_Comissioning[2],
                   HMI_EStop := "PLC_HMI - HMI 2 Estop",
                   HMI_Profinet_Error := "PLC_HMI - Profinet_Error_HMI 2",
                   Local_Mode := "HMI_2_Local_Mode",
                   HMI_Estop_Pressed_1 => #HMI_2_Estop_Pressed_1,
                   HMI_Estop_Pressed_2 => #HMI_2_Estop_Pressed_2,
                   HMI_Estop_Pressed_3 => #HMI_2_Estop_Pressed_3,
                   HMI_Estop_Pressed_4 => #HMI_2_Estop_Pressed_4,
                   HMI_Estop_Pressed_5 => #HMI_2_Estop_Pressed_5,
                   Reset_Comissioning_1 => #HMI_2_Reset_Comiss_1,
                   Reset_Comissioning_2 => #HMI_2_Reset_Comiss_2,
                   Reset_Comissioning_3 => #HMI_2_Reset_Comiss_3,
                   Reset_Comissioning_4 => #HMI_2_Reset_Comiss_4,
                   Reset_Comissioning_5 => #HMI_2_Reset_Comiss_5);
END_REGION

REGION Network 4: Remote Panel 1
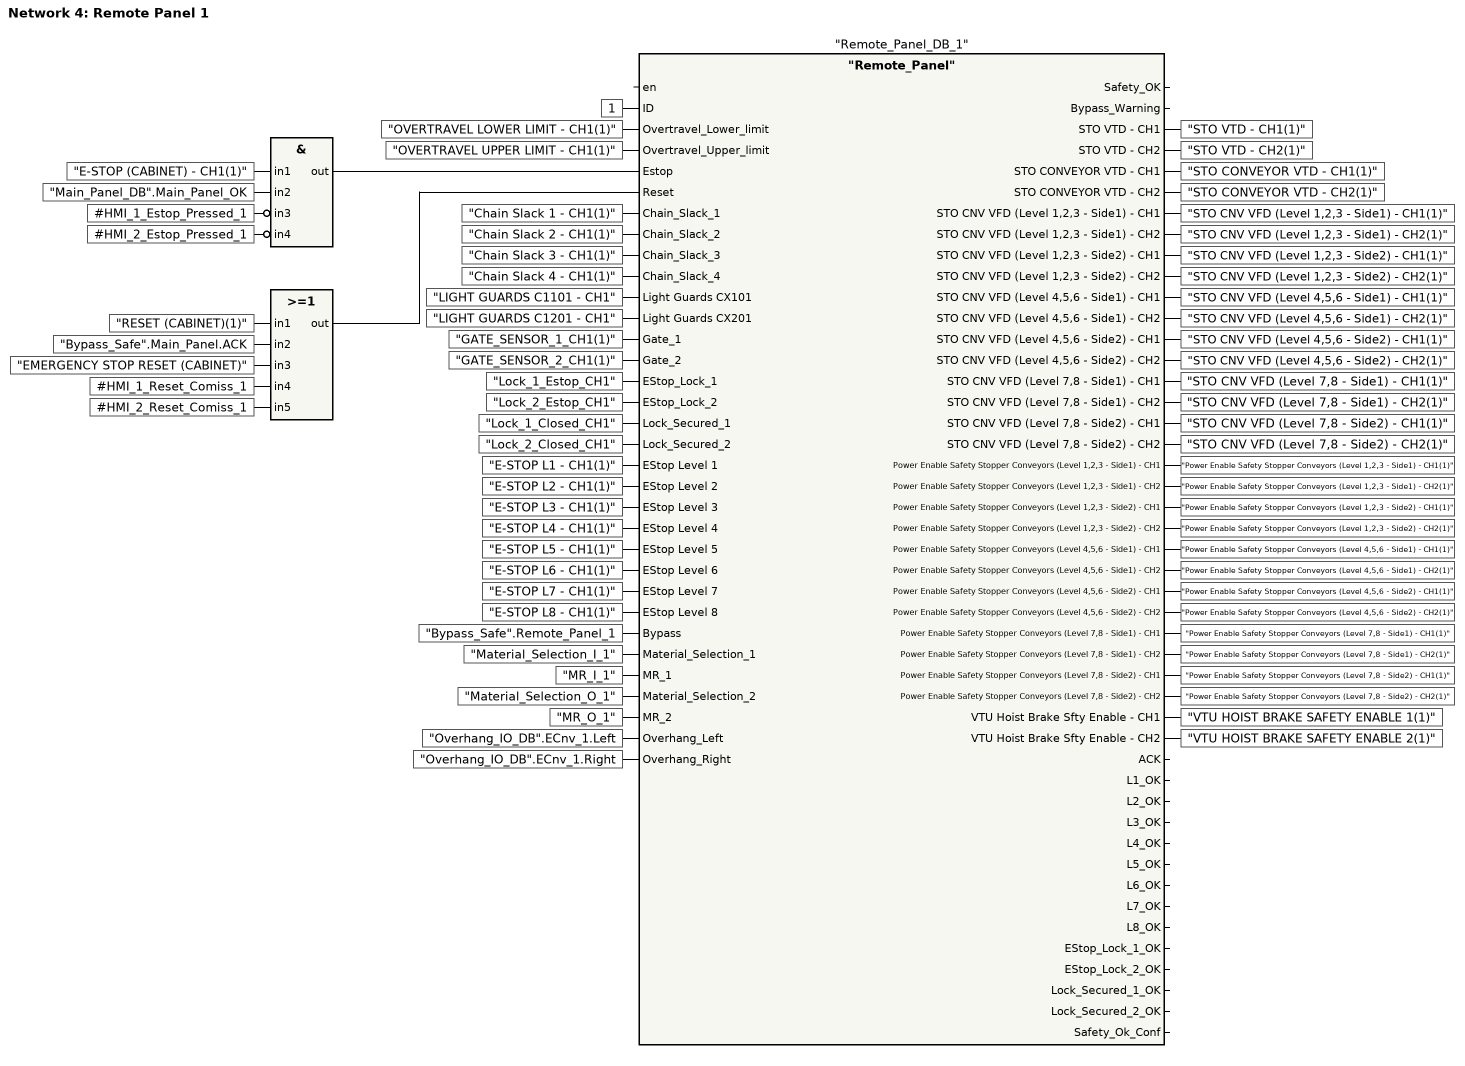
   "Remote_Panel_DB_1"(ID := 1,   // "Remote_Panel"
                       Overtravel_Lower_limit := "OVERTRAVEL LOWER LIMIT - CH1(1)",
                       Overtravel_Upper_limit := "OVERTRAVEL UPPER LIMIT - CH1(1)",
                       Estop := "E-STOP (CABINET) - CH1(1)" AND "Main_Panel_DB".Main_Panel_OK AND NOT #HMI_1_Estop_Pressed_1 AND NOT #HMI_2_Estop_Pressed_1,
                       Reset := "RESET (CABINET)(1)" OR "Bypass_Safe".Main_Panel.ACK OR "EMERGENCY STOP RESET (CABINET)" OR #HMI_1_Reset_Comiss_1 OR #HMI_2_Reset_Comiss_1,
                       Chain_Slack_1 := "Chain Slack 1 - CH1(1)",
                       Chain_Slack_2 := "Chain Slack 2 - CH1(1)",
                       Chain_Slack_3 := "Chain Slack 3 - CH1(1)",
                       Chain_Slack_4 := "Chain Slack 4 - CH1(1)",
                       "Light Guards CX101" := "LIGHT GUARDS C1101 - CH1",
                       "Light Guards CX201" := "LIGHT GUARDS C1201 - CH1",
                       Gate_1 := "GATE_SENSOR_1_CH1(1)",
                       Gate_2 := "GATE_SENSOR_2_CH1(1)",
                       EStop_Lock_1 := "Lock_1_Estop_CH1",
                       EStop_Lock_2 := "Lock_2_Estop_CH1",
                       Lock_Secured_1 := "Lock_1_Closed_CH1",
                       Lock_Secured_2 := "Lock_2_Closed_CH1",
                       "EStop Level 1" := "E-STOP L1 - CH1(1)",
                       "EStop Level 2" := "E-STOP L2 - CH1(1)",
                       "EStop Level 3" := "E-STOP L3 - CH1(1)",
                       "EStop Level 4" := "E-STOP L4 - CH1(1)",
                       "EStop Level 5" := "E-STOP L5 - CH1(1)",
                       "EStop Level 6" := "E-STOP L6 - CH1(1)",
                       "EStop Level 7" := "E-STOP L7 - CH1(1)",
                       "EStop Level 8" := "E-STOP L8 - CH1(1)",
                       Bypass := "Bypass_Safe".Remote_Panel_1,
                       Material_Selection_1 := "Material_Selection_I_1",
                       MR_1 := "MR_I_1",
                       Material_Selection_2 := "Material_Selection_O_1",
                       MR_2 := "MR_O_1",
                       Overhang_Left := "Overhang_IO_DB".ECnv_1.Left,
                       Overhang_Right := "Overhang_IO_DB".ECnv_1.Right,
                       "STO VTD - CH1" => "STO VTD - CH1(1)",
                       "STO VTD - CH2" => "STO VTD - CH2(1)",
                       "STO CONVEYOR VTD - CH1" => "STO CONVEYOR VTD - CH1(1)",
                       "STO CONVEYOR VTD - CH2" => "STO CONVEYOR VTD - CH2(1)",
                       "STO CNV VFD (Level 1,2,3 - Side1) - CH1" => "STO CNV VFD (Level 1,2,3 - Side1) - CH1(1)",
                       "STO CNV VFD (Level 1,2,3 - Side1) - CH2" => "STO CNV VFD (Level 1,2,3 - Side1) - CH2(1)",
                       "STO CNV VFD (Level 1,2,3 - Side2) - CH1" => "STO CNV VFD (Level 1,2,3 - Side2) - CH1(1)",
                       "STO CNV VFD (Level 1,2,3 - Side2) - CH2" => "STO CNV VFD (Level 1,2,3 - Side2) - CH2(1)",
                       "STO CNV VFD (Level 4,5,6 - Side1) - CH1" => "STO CNV VFD (Level 4,5,6 - Side1) - CH1(1)",
                       "STO CNV VFD (Level 4,5,6 - Side1) - CH2" => "STO CNV VFD (Level 4,5,6 - Side1) - CH2(1)",
                       "STO CNV VFD (Level 4,5,6 - Side2) - CH1" => "STO CNV VFD (Level 4,5,6 - Side2) - CH1(1)",
                       "STO CNV VFD (Level 4,5,6 - Side2) - CH2" => "STO CNV VFD (Level 4,5,6 - Side2) - CH2(1)",
                       "STO CNV VFD (Level 7,8 - Side1) - CH1" => "STO CNV VFD (Level 7,8 - Side1) - CH1(1)",
                       "STO CNV VFD (Level 7,8 - Side1) - CH2" => "STO CNV VFD (Level 7,8 - Side1) - CH2(1)",
                       "STO CNV VFD (Level 7,8 - Side2) - CH1" => "STO CNV VFD (Level 7,8 - Side2) - CH1(1)",
                       "STO CNV VFD (Level 7,8 - Side2) - CH2" => "STO CNV VFD (Level 7,8 - Side2) - CH2(1)",
                       "Power Enable Safety Stopper Conveyors (Level 1,2,3 - Side1) - CH1" => "Power Enable Safety Stopper Conveyors (Level 1,2,3 - Side1) - CH1(1)",
                       "Power Enable Safety Stopper Conveyors (Level 1,2,3 - Side1) - CH2" => "Power Enable Safety Stopper Conveyors (Level 1,2,3 - Side1) - CH2(1)",
                       "Power Enable Safety Stopper Conveyors (Level 1,2,3 - Side2) - CH1" => "Power Enable Safety Stopper Conveyors (Level 1,2,3 - Side2) - CH1(1)",
                       "Power Enable Safety Stopper Conveyors (Level 1,2,3 - Side2) - CH2" => "Power Enable Safety Stopper Conveyors (Level 1,2,3 - Side2) - CH2(1)",
                       "Power Enable Safety Stopper Conveyors (Level 4,5,6 - Side1) - CH1" => "Power Enable Safety Stopper Conveyors (Level 4,5,6 - Side1) - CH1(1)",
                       "Power Enable Safety Stopper Conveyors (Level 4,5,6 - Side1) - CH2" => "Power Enable Safety Stopper Conveyors (Level 4,5,6 - Side1) - CH2(1)",
                       "Power Enable Safety Stopper Conveyors (Level 4,5,6 - Side2) - CH1" => "Power Enable Safety Stopper Conveyors (Level 4,5,6 - Side2) - CH1(1)",
                       "Power Enable Safety Stopper Conveyors (Level 4,5,6 - Side2) - CH2" => "Power Enable Safety Stopper Conveyors (Level 4,5,6 - Side2) - CH2(1)",
                       "Power Enable Safety Stopper Conveyors (Level 7,8 - Side1) - CH1" => "Power Enable Safety Stopper Conveyors (Level 7,8 - Side1) - CH1(1)",
                       "Power Enable Safety Stopper Conveyors (Level 7,8 - Side1) - CH2" => "Power Enable Safety Stopper Conveyors (Level 7,8 - Side1) - CH2(1)",
                       "Power Enable Safety Stopper Conveyors (Level 7,8 - Side2) - CH1" => "Power Enable Safety Stopper Conveyors (Level 7,8 - Side2) - CH1(1)",
                       "Power Enable Safety Stopper Conveyors (Level 7,8 - Side2) - CH2" => "Power Enable Safety Stopper Conveyors (Level 7,8 - Side2) - CH2(1)",
                       "VTU Hoist Brake Sfty Enable - CH1" => "VTU HOIST BRAKE SAFETY ENABLE 1(1)",
                       "VTU Hoist Brake Sfty Enable - CH2" => "VTU HOIST BRAKE SAFETY ENABLE 2(1)");
END_REGION

REGION Network 5: Remote Panel 2
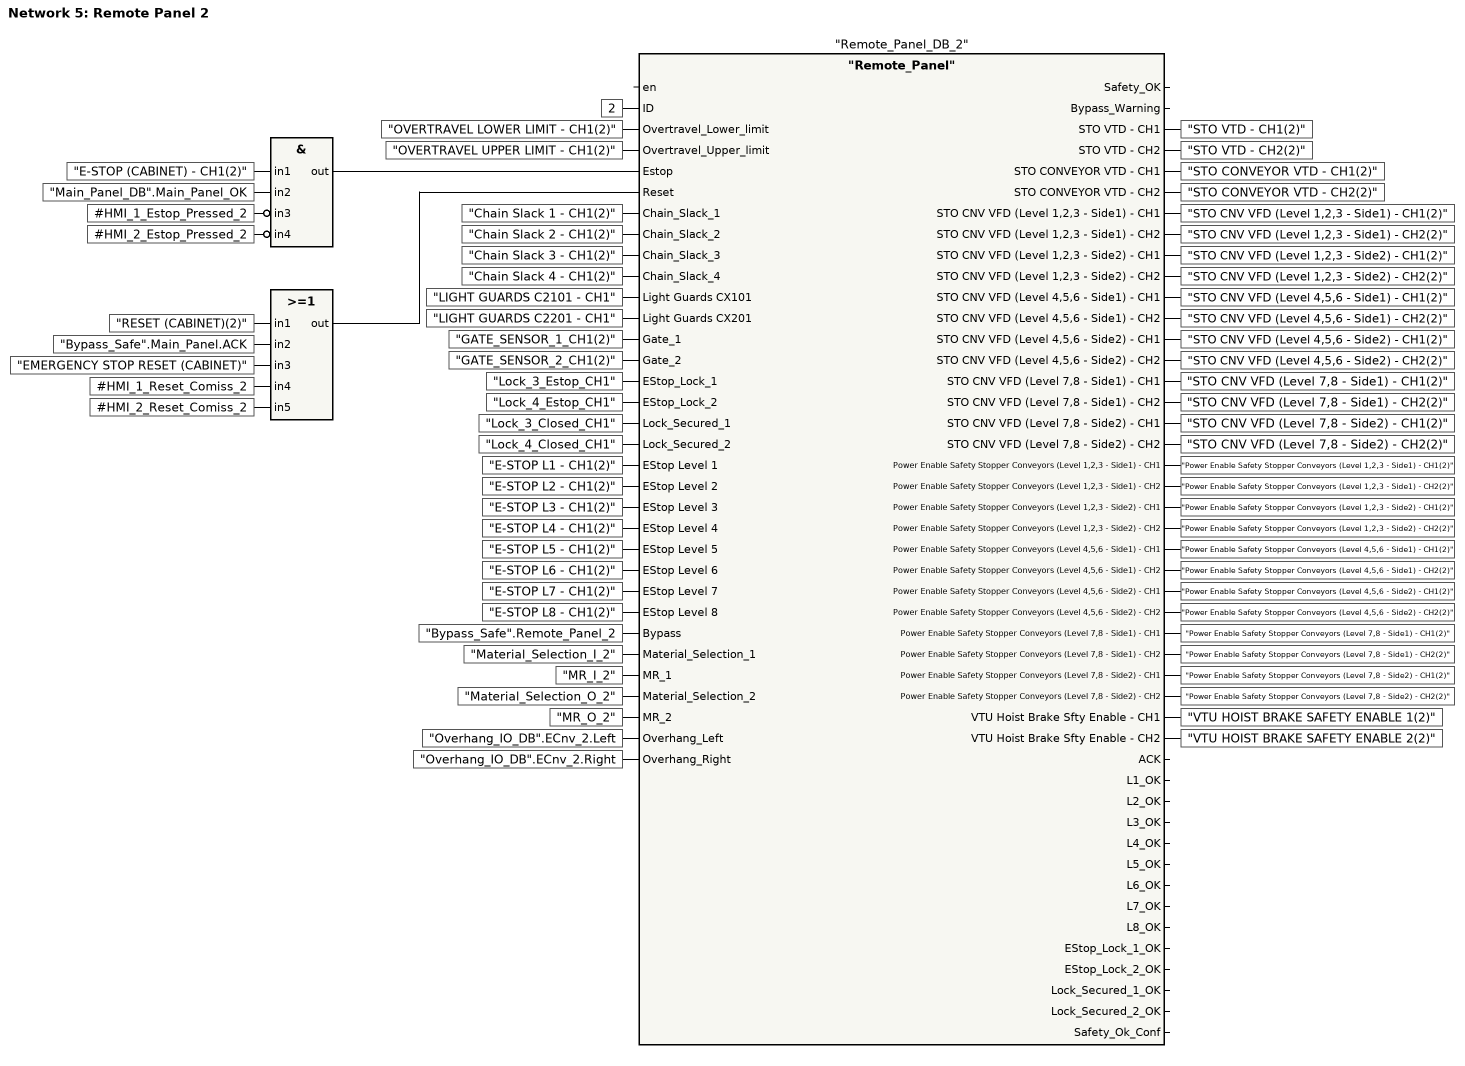
   "Remote_Panel_DB_2"(ID := 2,   // "Remote_Panel"
                       Overtravel_Lower_limit := "OVERTRAVEL LOWER LIMIT - CH1(2)",
                       Overtravel_Upper_limit := "OVERTRAVEL UPPER LIMIT - CH1(2)",
                       Estop := "E-STOP (CABINET) - CH1(2)" AND "Main_Panel_DB".Main_Panel_OK AND NOT #HMI_1_Estop_Pressed_2 AND NOT #HMI_2_Estop_Pressed_2,
                       Reset := "RESET (CABINET)(2)" OR "Bypass_Safe".Main_Panel.ACK OR "EMERGENCY STOP RESET (CABINET)" OR #HMI_1_Reset_Comiss_2 OR #HMI_2_Reset_Comiss_2,
                       Chain_Slack_1 := "Chain Slack 1 - CH1(2)",
                       Chain_Slack_2 := "Chain Slack 2 - CH1(2)",
                       Chain_Slack_3 := "Chain Slack 3 - CH1(2)",
                       Chain_Slack_4 := "Chain Slack 4 - CH1(2)",
                       "Light Guards CX101" := "LIGHT GUARDS C2101 - CH1",
                       "Light Guards CX201" := "LIGHT GUARDS C2201 - CH1",
                       Gate_1 := "GATE_SENSOR_1_CH1(2)",
                       Gate_2 := "GATE_SENSOR_2_CH1(2)",
                       EStop_Lock_1 := "Lock_3_Estop_CH1",
                       EStop_Lock_2 := "Lock_4_Estop_CH1",
                       Lock_Secured_1 := "Lock_3_Closed_CH1",
                       Lock_Secured_2 := "Lock_4_Closed_CH1",
                       "EStop Level 1" := "E-STOP L1 - CH1(2)",
                       "EStop Level 2" := "E-STOP L2 - CH1(2)",
                       "EStop Level 3" := "E-STOP L3 - CH1(2)",
                       "EStop Level 4" := "E-STOP L4 - CH1(2)",
                       "EStop Level 5" := "E-STOP L5 - CH1(2)",
                       "EStop Level 6" := "E-STOP L6 - CH1(2)",
                       "EStop Level 7" := "E-STOP L7 - CH1(2)",
                       "EStop Level 8" := "E-STOP L8 - CH1(2)",
                       Bypass := "Bypass_Safe".Remote_Panel_2,
                       Material_Selection_1 := "Material_Selection_I_2",
                       MR_1 := "MR_I_2",
                       Material_Selection_2 := "Material_Selection_O_2",
                       MR_2 := "MR_O_2",
                       Overhang_Left := "Overhang_IO_DB".ECnv_2.Left,
                       Overhang_Right := "Overhang_IO_DB".ECnv_2.Right,
                       "STO VTD - CH1" => "STO VTD - CH1(2)",
                       "STO VTD - CH2" => "STO VTD - CH2(2)",
                       "STO CONVEYOR VTD - CH1" => "STO CONVEYOR VTD - CH1(2)",
                       "STO CONVEYOR VTD - CH2" => "STO CONVEYOR VTD - CH2(2)",
                       "STO CNV VFD (Level 1,2,3 - Side1) - CH1" => "STO CNV VFD (Level 1,2,3 - Side1) - CH1(2)",
                       "STO CNV VFD (Level 1,2,3 - Side1) - CH2" => "STO CNV VFD (Level 1,2,3 - Side1) - CH2(2)",
                       "STO CNV VFD (Level 1,2,3 - Side2) - CH1" => "STO CNV VFD (Level 1,2,3 - Side2) - CH1(2)",
                       "STO CNV VFD (Level 1,2,3 - Side2) - CH2" => "STO CNV VFD (Level 1,2,3 - Side2) - CH2(2)",
                       "STO CNV VFD (Level 4,5,6 - Side1) - CH1" => "STO CNV VFD (Level 4,5,6 - Side1) - CH1(2)",
                       "STO CNV VFD (Level 4,5,6 - Side1) - CH2" => "STO CNV VFD (Level 4,5,6 - Side1) - CH2(2)",
                       "STO CNV VFD (Level 4,5,6 - Side2) - CH1" => "STO CNV VFD (Level 4,5,6 - Side2) - CH1(2)",
                       "STO CNV VFD (Level 4,5,6 - Side2) - CH2" => "STO CNV VFD (Level 4,5,6 - Side2) - CH2(2)",
                       "STO CNV VFD (Level 7,8 - Side1) - CH1" => "STO CNV VFD (Level 7,8 - Side1) - CH1(2)",
                       "STO CNV VFD (Level 7,8 - Side1) - CH2" => "STO CNV VFD (Level 7,8 - Side1) - CH2(2)",
                       "STO CNV VFD (Level 7,8 - Side2) - CH1" => "STO CNV VFD (Level 7,8 - Side2) - CH1(2)",
                       "STO CNV VFD (Level 7,8 - Side2) - CH2" => "STO CNV VFD (Level 7,8 - Side2) - CH2(2)",
                       "Power Enable Safety Stopper Conveyors (Level 1,2,3 - Side1) - CH1" => "Power Enable Safety Stopper Conveyors (Level 1,2,3 - Side1) - CH1(2)",
                       "Power Enable Safety Stopper Conveyors (Level 1,2,3 - Side1) - CH2" => "Power Enable Safety Stopper Conveyors (Level 1,2,3 - Side1) - CH2(2)",
                       "Power Enable Safety Stopper Conveyors (Level 1,2,3 - Side2) - CH1" => "Power Enable Safety Stopper Conveyors (Level 1,2,3 - Side2) - CH1(2)",
                       "Power Enable Safety Stopper Conveyors (Level 1,2,3 - Side2) - CH2" => "Power Enable Safety Stopper Conveyors (Level 1,2,3 - Side2) - CH2(2)",
                       "Power Enable Safety Stopper Conveyors (Level 4,5,6 - Side1) - CH1" => "Power Enable Safety Stopper Conveyors (Level 4,5,6 - Side1) - CH1(2)",
                       "Power Enable Safety Stopper Conveyors (Level 4,5,6 - Side1) - CH2" => "Power Enable Safety Stopper Conveyors (Level 4,5,6 - Side1) - CH2(2)",
                       "Power Enable Safety Stopper Conveyors (Level 4,5,6 - Side2) - CH1" => "Power Enable Safety Stopper Conveyors (Level 4,5,6 - Side2) - CH1(2)",
                       "Power Enable Safety Stopper Conveyors (Level 4,5,6 - Side2) - CH2" => "Power Enable Safety Stopper Conveyors (Level 4,5,6 - Side2) - CH2(2)",
                       "Power Enable Safety Stopper Conveyors (Level 7,8 - Side1) - CH1" => "Power Enable Safety Stopper Conveyors (Level 7,8 - Side1) - CH1(2)",
                       "Power Enable Safety Stopper Conveyors (Level 7,8 - Side1) - CH2" => "Power Enable Safety Stopper Conveyors (Level 7,8 - Side1) - CH2(2)",
                       "Power Enable Safety Stopper Conveyors (Level 7,8 - Side2) - CH1" => "Power Enable Safety Stopper Conveyors (Level 7,8 - Side2) - CH1(2)",
                       "Power Enable Safety Stopper Conveyors (Level 7,8 - Side2) - CH2" => "Power Enable Safety Stopper Conveyors (Level 7,8 - Side2) - CH2(2)",
                       "VTU Hoist Brake Sfty Enable - CH1" => "VTU HOIST BRAKE SAFETY ENABLE 1(2)",
                       "VTU Hoist Brake Sfty Enable - CH2" => "VTU HOIST BRAKE SAFETY ENABLE 2(2)");
END_REGION

REGION Network 6: Remote Panel 3
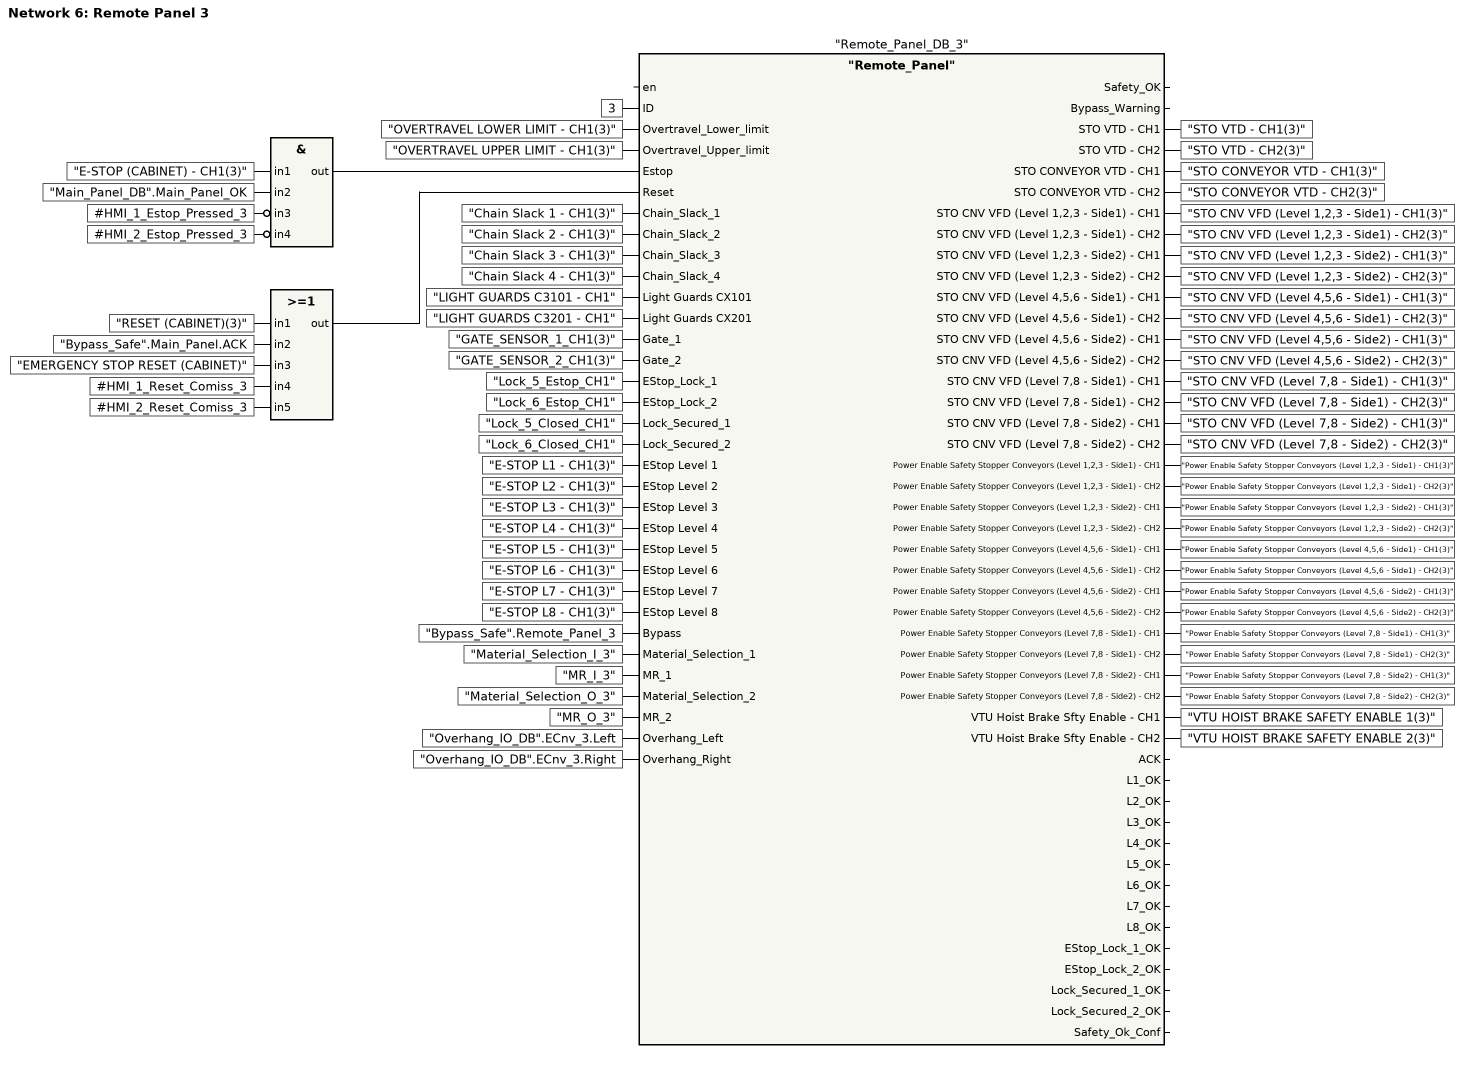
   "Remote_Panel_DB_3"(ID := 3,   // "Remote_Panel"
                       Overtravel_Lower_limit := "OVERTRAVEL LOWER LIMIT - CH1(3)",
                       Overtravel_Upper_limit := "OVERTRAVEL UPPER LIMIT - CH1(3)",
                       Estop := "E-STOP (CABINET) - CH1(3)" AND "Main_Panel_DB".Main_Panel_OK AND NOT #HMI_1_Estop_Pressed_3 AND NOT #HMI_2_Estop_Pressed_3,
                       Reset := "RESET (CABINET)(3)" OR "Bypass_Safe".Main_Panel.ACK OR "EMERGENCY STOP RESET (CABINET)" OR #HMI_1_Reset_Comiss_3 OR #HMI_2_Reset_Comiss_3,
                       Chain_Slack_1 := "Chain Slack 1 - CH1(3)",
                       Chain_Slack_2 := "Chain Slack 2 - CH1(3)",
                       Chain_Slack_3 := "Chain Slack 3 - CH1(3)",
                       Chain_Slack_4 := "Chain Slack 4 - CH1(3)",
                       "Light Guards CX101" := "LIGHT GUARDS C3101 - CH1",
                       "Light Guards CX201" := "LIGHT GUARDS C3201 - CH1",
                       Gate_1 := "GATE_SENSOR_1_CH1(3)",
                       Gate_2 := "GATE_SENSOR_2_CH1(3)",
                       EStop_Lock_1 := "Lock_5_Estop_CH1",
                       EStop_Lock_2 := "Lock_6_Estop_CH1",
                       Lock_Secured_1 := "Lock_5_Closed_CH1",
                       Lock_Secured_2 := "Lock_6_Closed_CH1",
                       "EStop Level 1" := "E-STOP L1 - CH1(3)",
                       "EStop Level 2" := "E-STOP L2 - CH1(3)",
                       "EStop Level 3" := "E-STOP L3 - CH1(3)",
                       "EStop Level 4" := "E-STOP L4 - CH1(3)",
                       "EStop Level 5" := "E-STOP L5 - CH1(3)",
                       "EStop Level 6" := "E-STOP L6 - CH1(3)",
                       "EStop Level 7" := "E-STOP L7 - CH1(3)",
                       "EStop Level 8" := "E-STOP L8 - CH1(3)",
                       Bypass := "Bypass_Safe".Remote_Panel_3,
                       Material_Selection_1 := "Material_Selection_I_3",
                       MR_1 := "MR_I_3",
                       Material_Selection_2 := "Material_Selection_O_3",
                       MR_2 := "MR_O_3",
                       Overhang_Left := "Overhang_IO_DB".ECnv_3.Left,
                       Overhang_Right := "Overhang_IO_DB".ECnv_3.Right,
                       "STO VTD - CH1" => "STO VTD - CH1(3)",
                       "STO VTD - CH2" => "STO VTD - CH2(3)",
                       "STO CONVEYOR VTD - CH1" => "STO CONVEYOR VTD - CH1(3)",
                       "STO CONVEYOR VTD - CH2" => "STO CONVEYOR VTD - CH2(3)",
                       "STO CNV VFD (Level 1,2,3 - Side1) - CH1" => "STO CNV VFD (Level 1,2,3 - Side1) - CH1(3)",
                       "STO CNV VFD (Level 1,2,3 - Side1) - CH2" => "STO CNV VFD (Level 1,2,3 - Side1) - CH2(3)",
                       "STO CNV VFD (Level 1,2,3 - Side2) - CH1" => "STO CNV VFD (Level 1,2,3 - Side2) - CH1(3)",
                       "STO CNV VFD (Level 1,2,3 - Side2) - CH2" => "STO CNV VFD (Level 1,2,3 - Side2) - CH2(3)",
                       "STO CNV VFD (Level 4,5,6 - Side1) - CH1" => "STO CNV VFD (Level 4,5,6 - Side1) - CH1(3)",
                       "STO CNV VFD (Level 4,5,6 - Side1) - CH2" => "STO CNV VFD (Level 4,5,6 - Side1) - CH2(3)",
                       "STO CNV VFD (Level 4,5,6 - Side2) - CH1" => "STO CNV VFD (Level 4,5,6 - Side2) - CH1(3)",
                       "STO CNV VFD (Level 4,5,6 - Side2) - CH2" => "STO CNV VFD (Level 4,5,6 - Side2) - CH2(3)",
                       "STO CNV VFD (Level 7,8 - Side1) - CH1" => "STO CNV VFD (Level 7,8 - Side1) - CH1(3)",
                       "STO CNV VFD (Level 7,8 - Side1) - CH2" => "STO CNV VFD (Level 7,8 - Side1) - CH2(3)",
                       "STO CNV VFD (Level 7,8 - Side2) - CH1" => "STO CNV VFD (Level 7,8 - Side2) - CH1(3)",
                       "STO CNV VFD (Level 7,8 - Side2) - CH2" => "STO CNV VFD (Level 7,8 - Side2) - CH2(3)",
                       "Power Enable Safety Stopper Conveyors (Level 1,2,3 - Side1) - CH1" => "Power Enable Safety Stopper Conveyors (Level 1,2,3 - Side1) - CH1(3)",
                       "Power Enable Safety Stopper Conveyors (Level 1,2,3 - Side1) - CH2" => "Power Enable Safety Stopper Conveyors (Level 1,2,3 - Side1) - CH2(3)",
                       "Power Enable Safety Stopper Conveyors (Level 1,2,3 - Side2) - CH1" => "Power Enable Safety Stopper Conveyors (Level 1,2,3 - Side2) - CH1(3)",
                       "Power Enable Safety Stopper Conveyors (Level 1,2,3 - Side2) - CH2" => "Power Enable Safety Stopper Conveyors (Level 1,2,3 - Side2) - CH2(3)",
                       "Power Enable Safety Stopper Conveyors (Level 4,5,6 - Side1) - CH1" => "Power Enable Safety Stopper Conveyors (Level 4,5,6 - Side1) - CH1(3)",
                       "Power Enable Safety Stopper Conveyors (Level 4,5,6 - Side1) - CH2" => "Power Enable Safety Stopper Conveyors (Level 4,5,6 - Side1) - CH2(3)",
                       "Power Enable Safety Stopper Conveyors (Level 4,5,6 - Side2) - CH1" => "Power Enable Safety Stopper Conveyors (Level 4,5,6 - Side2) - CH1(3)",
                       "Power Enable Safety Stopper Conveyors (Level 4,5,6 - Side2) - CH2" => "Power Enable Safety Stopper Conveyors (Level 4,5,6 - Side2) - CH2(3)",
                       "Power Enable Safety Stopper Conveyors (Level 7,8 - Side1) - CH1" => "Power Enable Safety Stopper Conveyors (Level 7,8 - Side1) - CH1(3)",
                       "Power Enable Safety Stopper Conveyors (Level 7,8 - Side1) - CH2" => "Power Enable Safety Stopper Conveyors (Level 7,8 - Side1) - CH2(3)",
                       "Power Enable Safety Stopper Conveyors (Level 7,8 - Side2) - CH1" => "Power Enable Safety Stopper Conveyors (Level 7,8 - Side2) - CH1(3)",
                       "Power Enable Safety Stopper Conveyors (Level 7,8 - Side2) - CH2" => "Power Enable Safety Stopper Conveyors (Level 7,8 - Side2) - CH2(3)",
                       "VTU Hoist Brake Sfty Enable - CH1" => "VTU HOIST BRAKE SAFETY ENABLE 1(3)",
                       "VTU Hoist Brake Sfty Enable - CH2" => "VTU HOIST BRAKE SAFETY ENABLE 2(3)");
END_REGION

REGION Network 7: Remote Panel 4
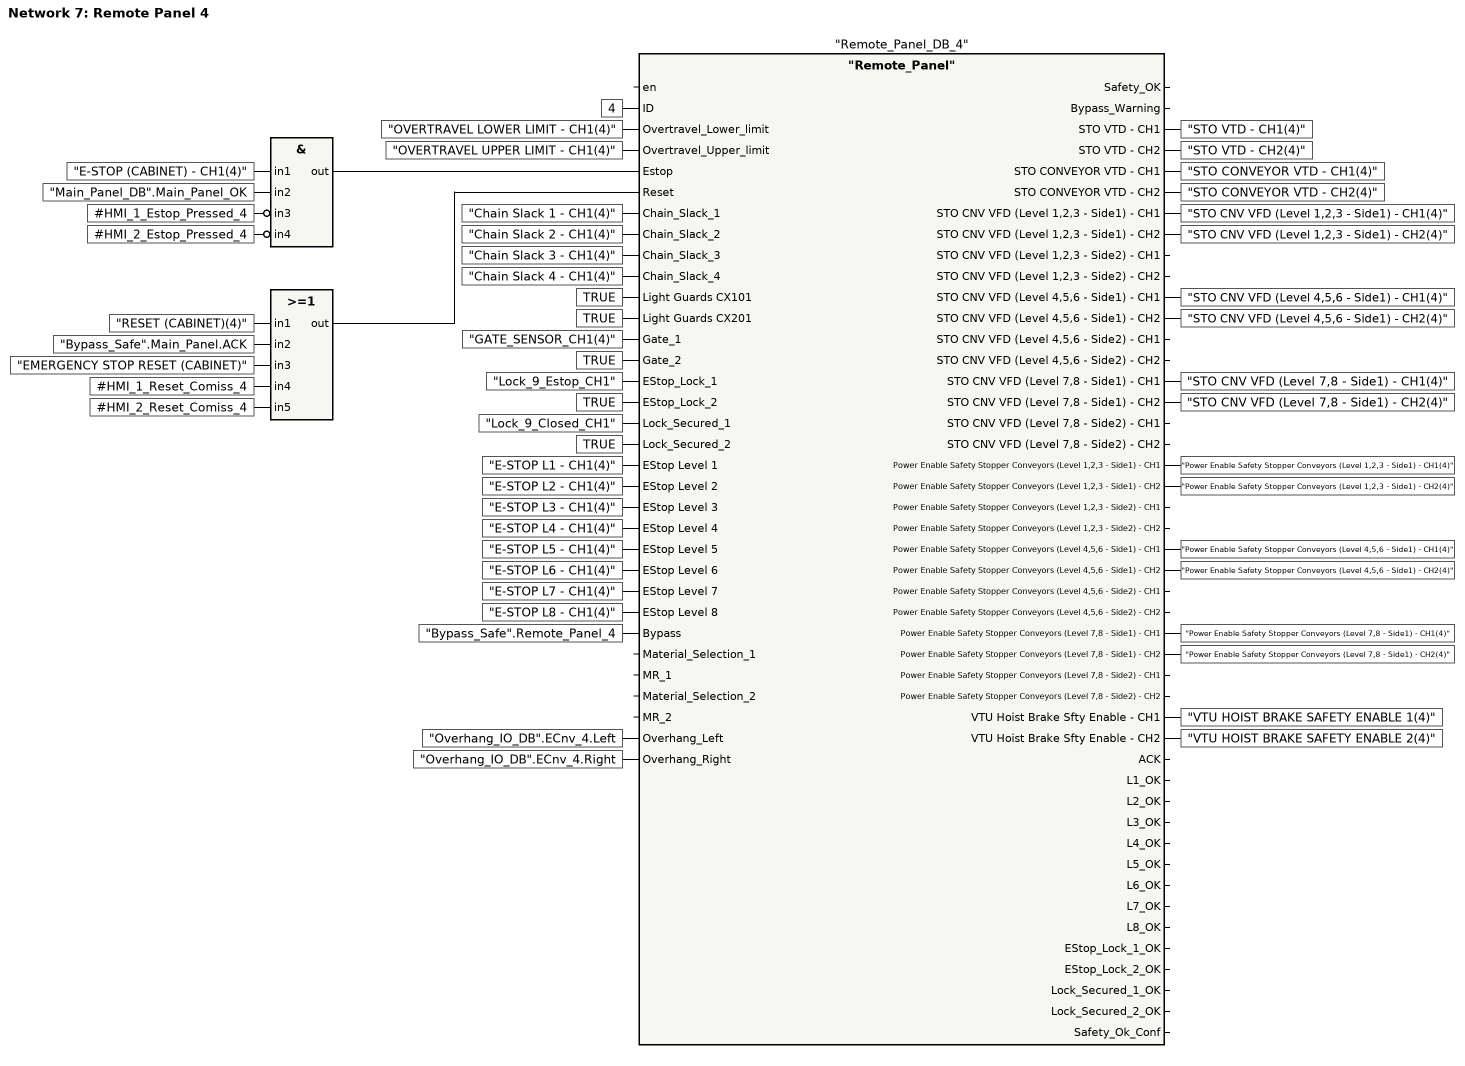
   "Remote_Panel_DB_4"(ID := 4,   // "Remote_Panel"
                       Overtravel_Lower_limit := "OVERTRAVEL LOWER LIMIT - CH1(4)",
                       Overtravel_Upper_limit := "OVERTRAVEL UPPER LIMIT - CH1(4)",
                       Estop := "E-STOP (CABINET) - CH1(4)" AND "Main_Panel_DB".Main_Panel_OK AND NOT #HMI_1_Estop_Pressed_4 AND NOT #HMI_2_Estop_Pressed_4,
                       Reset := "RESET (CABINET)(4)" OR "Bypass_Safe".Main_Panel.ACK OR "EMERGENCY STOP RESET (CABINET)" OR #HMI_1_Reset_Comiss_4 OR #HMI_2_Reset_Comiss_4,
                       Chain_Slack_1 := "Chain Slack 1 - CH1(4)",
                       Chain_Slack_2 := "Chain Slack 2 - CH1(4)",
                       Chain_Slack_3 := "Chain Slack 3 - CH1(4)",
                       Chain_Slack_4 := "Chain Slack 4 - CH1(4)",
                       "Light Guards CX101" := TRUE,
                       "Light Guards CX201" := TRUE,
                       Gate_1 := "GATE_SENSOR_CH1(4)",
                       Gate_2 := TRUE,
                       EStop_Lock_1 := "Lock_9_Estop_CH1",
                       EStop_Lock_2 := TRUE,
                       Lock_Secured_1 := "Lock_9_Closed_CH1",
                       Lock_Secured_2 := TRUE,
                       "EStop Level 1" := "E-STOP L1 - CH1(4)",
                       "EStop Level 2" := "E-STOP L2 - CH1(4)",
                       "EStop Level 3" := "E-STOP L3 - CH1(4)",
                       "EStop Level 4" := "E-STOP L4 - CH1(4)",
                       "EStop Level 5" := "E-STOP L5 - CH1(4)",
                       "EStop Level 6" := "E-STOP L6 - CH1(4)",
                       "EStop Level 7" := "E-STOP L7 - CH1(4)",
                       "EStop Level 8" := "E-STOP L8 - CH1(4)",
                       Bypass := "Bypass_Safe".Remote_Panel_4,
                       Overhang_Left := "Overhang_IO_DB".ECnv_4.Left,
                       Overhang_Right := "Overhang_IO_DB".ECnv_4.Right,
                       "STO VTD - CH1" => "STO VTD - CH1(4)",
                       "STO VTD - CH2" => "STO VTD - CH2(4)",
                       "STO CONVEYOR VTD - CH1" => "STO CONVEYOR VTD - CH1(4)",
                       "STO CONVEYOR VTD - CH2" => "STO CONVEYOR VTD - CH2(4)",
                       "STO CNV VFD (Level 1,2,3 - Side1) - CH1" => "STO CNV VFD (Level 1,2,3 - Side1) - CH1(4)",
                       "STO CNV VFD (Level 1,2,3 - Side1) - CH2" => "STO CNV VFD (Level 1,2,3 - Side1) - CH2(4)",
                       "STO CNV VFD (Level 4,5,6 - Side1) - CH1" => "STO CNV VFD (Level 4,5,6 - Side1) - CH1(4)",
                       "STO CNV VFD (Level 4,5,6 - Side1) - CH2" => "STO CNV VFD (Level 4,5,6 - Side1) - CH2(4)",
                       "STO CNV VFD (Level 7,8 - Side1) - CH1" => "STO CNV VFD (Level 7,8 - Side1) - CH1(4)",
                       "STO CNV VFD (Level 7,8 - Side1) - CH2" => "STO CNV VFD (Level 7,8 - Side1) - CH2(4)",
                       "Power Enable Safety Stopper Conveyors (Level 1,2,3 - Side1) - CH1" => "Power Enable Safety Stopper Conveyors (Level 1,2,3 - Side1) - CH1(4)",
                       "Power Enable Safety Stopper Conveyors (Level 1,2,3 - Side1) - CH2" => "Power Enable Safety Stopper Conveyors (Level 1,2,3 - Side1) - CH2(4)",
                       "Power Enable Safety Stopper Conveyors (Level 4,5,6 - Side1) - CH1" => "Power Enable Safety Stopper Conveyors (Level 4,5,6 - Side1) - CH1(4)",
                       "Power Enable Safety Stopper Conveyors (Level 4,5,6 - Side1) - CH2" => "Power Enable Safety Stopper Conveyors (Level 4,5,6 - Side1) - CH2(4)",
                       "Power Enable Safety Stopper Conveyors (Level 7,8 - Side1) - CH1" => "Power Enable Safety Stopper Conveyors (Level 7,8 - Side1) - CH1(4)",
                       "Power Enable Safety Stopper Conveyors (Level 7,8 - Side1) - CH2" => "Power Enable Safety Stopper Conveyors (Level 7,8 - Side1) - CH2(4)",
                       "VTU Hoist Brake Sfty Enable - CH1" => "VTU HOIST BRAKE SAFETY ENABLE 1(4)",
                       "VTU Hoist Brake Sfty Enable - CH2" => "VTU HOIST BRAKE SAFETY ENABLE 2(4)");
END_REGION

REGION Network 8: Remote Panel 5
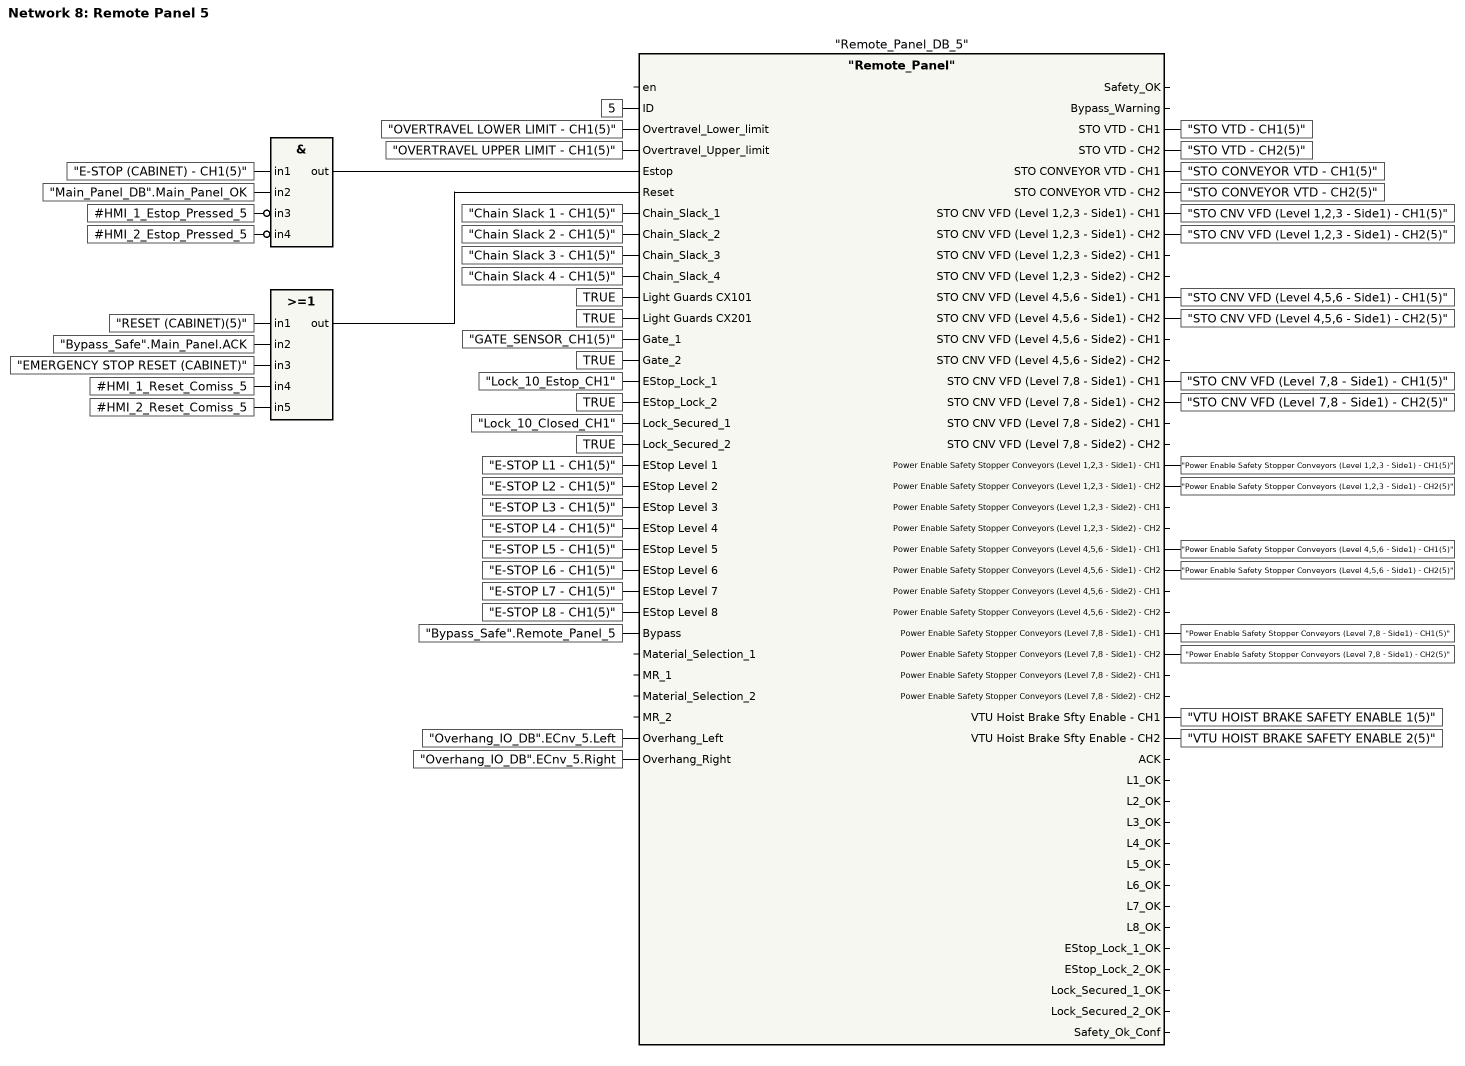
   "Remote_Panel_DB_5"(ID := 5,   // "Remote_Panel"
                       Overtravel_Lower_limit := "OVERTRAVEL LOWER LIMIT - CH1(5)",
                       Overtravel_Upper_limit := "OVERTRAVEL UPPER LIMIT - CH1(5)",
                       Estop := "E-STOP (CABINET) - CH1(5)" AND "Main_Panel_DB".Main_Panel_OK AND NOT #HMI_1_Estop_Pressed_5 AND NOT #HMI_2_Estop_Pressed_5,
                       Reset := "RESET (CABINET)(5)" OR "Bypass_Safe".Main_Panel.ACK OR "EMERGENCY STOP RESET (CABINET)" OR #HMI_1_Reset_Comiss_5 OR #HMI_2_Reset_Comiss_5,
                       Chain_Slack_1 := "Chain Slack 1 - CH1(5)",
                       Chain_Slack_2 := "Chain Slack 2 - CH1(5)",
                       Chain_Slack_3 := "Chain Slack 3 - CH1(5)",
                       Chain_Slack_4 := "Chain Slack 4 - CH1(5)",
                       "Light Guards CX101" := TRUE,
                       "Light Guards CX201" := TRUE,
                       Gate_1 := "GATE_SENSOR_CH1(5)",
                       Gate_2 := TRUE,
                       EStop_Lock_1 := "Lock_10_Estop_CH1",
                       EStop_Lock_2 := TRUE,
                       Lock_Secured_1 := "Lock_10_Closed_CH1",
                       Lock_Secured_2 := TRUE,
                       "EStop Level 1" := "E-STOP L1 - CH1(5)",
                       "EStop Level 2" := "E-STOP L2 - CH1(5)",
                       "EStop Level 3" := "E-STOP L3 - CH1(5)",
                       "EStop Level 4" := "E-STOP L4 - CH1(5)",
                       "EStop Level 5" := "E-STOP L5 - CH1(5)",
                       "EStop Level 6" := "E-STOP L6 - CH1(5)",
                       "EStop Level 7" := "E-STOP L7 - CH1(5)",
                       "EStop Level 8" := "E-STOP L8 - CH1(5)",
                       Bypass := "Bypass_Safe".Remote_Panel_5,
                       Overhang_Left := "Overhang_IO_DB".ECnv_5.Left,
                       Overhang_Right := "Overhang_IO_DB".ECnv_5.Right,
                       "STO VTD - CH1" => "STO VTD - CH1(5)",
                       "STO VTD - CH2" => "STO VTD - CH2(5)",
                       "STO CONVEYOR VTD - CH1" => "STO CONVEYOR VTD - CH1(5)",
                       "STO CONVEYOR VTD - CH2" => "STO CONVEYOR VTD - CH2(5)",
                       "STO CNV VFD (Level 1,2,3 - Side1) - CH1" => "STO CNV VFD (Level 1,2,3 - Side1) - CH1(5)",
                       "STO CNV VFD (Level 1,2,3 - Side1) - CH2" => "STO CNV VFD (Level 1,2,3 - Side1) - CH2(5)",
                       "STO CNV VFD (Level 4,5,6 - Side1) - CH1" => "STO CNV VFD (Level 4,5,6 - Side1) - CH1(5)",
                       "STO CNV VFD (Level 4,5,6 - Side1) - CH2" => "STO CNV VFD (Level 4,5,6 - Side1) - CH2(5)",
                       "STO CNV VFD (Level 7,8 - Side1) - CH1" => "STO CNV VFD (Level 7,8 - Side1) - CH1(5)",
                       "STO CNV VFD (Level 7,8 - Side1) - CH2" => "STO CNV VFD (Level 7,8 - Side1) - CH2(5)",
                       "Power Enable Safety Stopper Conveyors (Level 1,2,3 - Side1) - CH1" => "Power Enable Safety Stopper Conveyors (Level 1,2,3 - Side1) - CH1(5)",
                       "Power Enable Safety Stopper Conveyors (Level 1,2,3 - Side1) - CH2" => "Power Enable Safety Stopper Conveyors (Level 1,2,3 - Side1) - CH2(5)",
                       "Power Enable Safety Stopper Conveyors (Level 4,5,6 - Side1) - CH1" => "Power Enable Safety Stopper Conveyors (Level 4,5,6 - Side1) - CH1(5)",
                       "Power Enable Safety Stopper Conveyors (Level 4,5,6 - Side1) - CH2" => "Power Enable Safety Stopper Conveyors (Level 4,5,6 - Side1) - CH2(5)",
                       "Power Enable Safety Stopper Conveyors (Level 7,8 - Side1) - CH1" => "Power Enable Safety Stopper Conveyors (Level 7,8 - Side1) - CH1(5)",
                       "Power Enable Safety Stopper Conveyors (Level 7,8 - Side1) - CH2" => "Power Enable Safety Stopper Conveyors (Level 7,8 - Side1) - CH2(5)",
                       "VTU Hoist Brake Sfty Enable - CH1" => "VTU HOIST BRAKE SAFETY ENABLE 1(5)",
                       "VTU Hoist Brake Sfty Enable - CH2" => "VTU HOIST BRAKE SAFETY ENABLE 2(5)");
END_REGION

REGION Network 9: ESTOP LEVEL PANELS
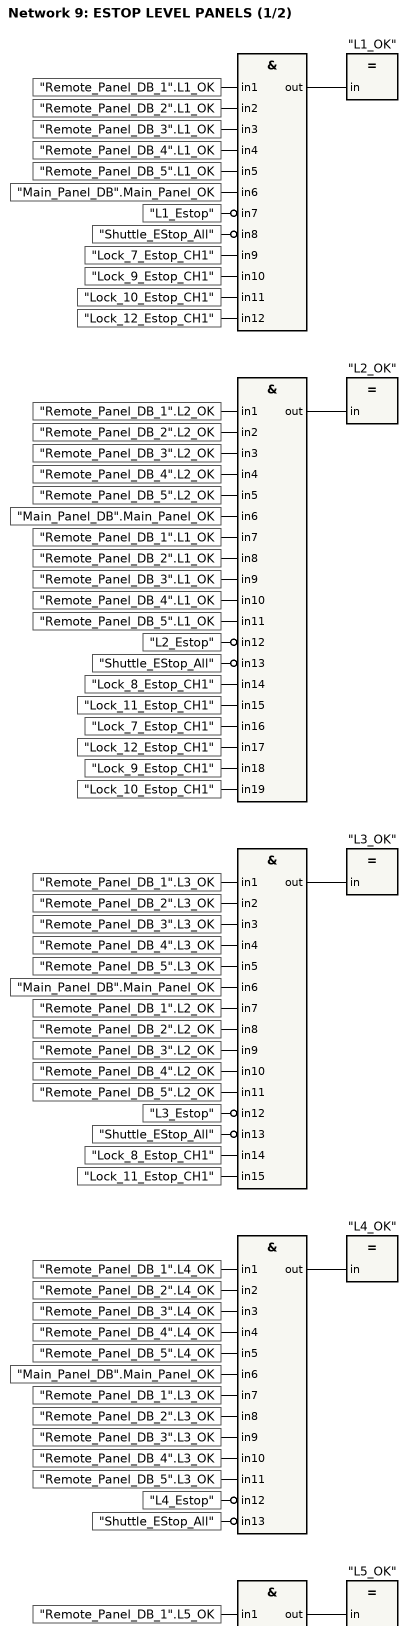
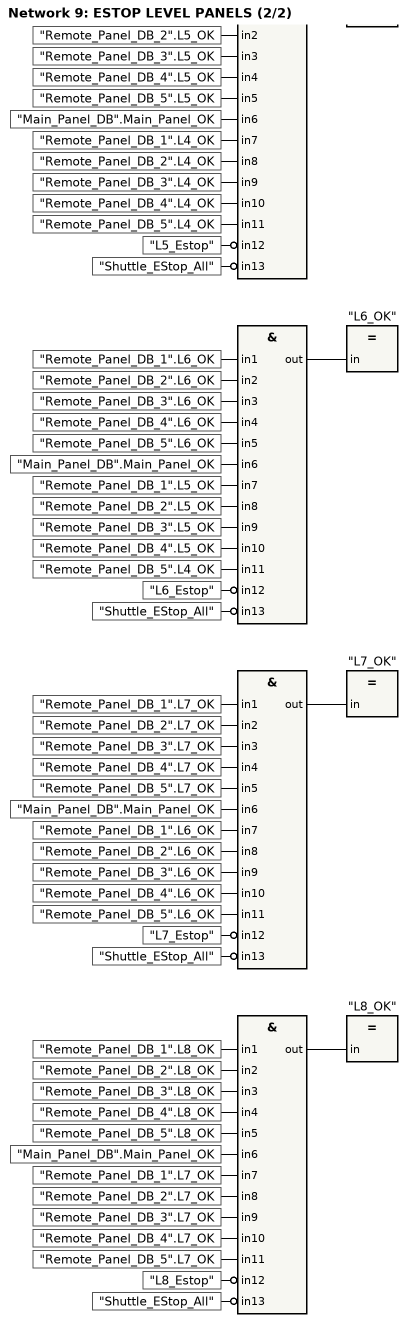
   "L1_OK" := "Remote_Panel_DB_1".L1_OK AND "Remote_Panel_DB_2".L1_OK AND "Remote_Panel_DB_3".L1_OK AND "Remote_Panel_DB_4".L1_OK AND "Remote_Panel_DB_5".L1_OK AND "Main_Panel_DB".Main_Panel_OK AND NOT "L1_Estop" AND NOT "Shuttle_EStop_All" AND "Lock_7_Estop_CH1" AND "Lock_9_Estop_CH1" AND "Lock_10_Estop_CH1" AND "Lock_12_Estop_CH1";
   "L2_OK" := "Remote_Panel_DB_1".L2_OK AND "Remote_Panel_DB_2".L2_OK AND "Remote_Panel_DB_3".L2_OK AND "Remote_Panel_DB_4".L2_OK AND "Remote_Panel_DB_5".L2_OK AND "Main_Panel_DB".Main_Panel_OK AND "Remote_Panel_DB_1".L1_OK AND "Remote_Panel_DB_2".L1_OK AND "Remote_Panel_DB_3".L1_OK AND "Remote_Panel_DB_4".L1_OK AND "Remote_Panel_DB_5".L1_OK AND NOT "L2_Estop" AND NOT "Shuttle_EStop_All" AND "Lock_8_Estop_CH1" AND "Lock_11_Estop_CH1" AND "Lock_7_Estop_CH1" AND "Lock_12_Estop_CH1" AND "Lock_9_Estop_CH1" AND "Lock_10_Estop_CH1";
   "L3_OK" := "Remote_Panel_DB_1".L3_OK AND "Remote_Panel_DB_2".L3_OK AND "Remote_Panel_DB_3".L3_OK AND "Remote_Panel_DB_4".L3_OK AND "Remote_Panel_DB_5".L3_OK AND "Main_Panel_DB".Main_Panel_OK AND "Remote_Panel_DB_1".L2_OK AND "Remote_Panel_DB_2".L2_OK AND "Remote_Panel_DB_3".L2_OK AND "Remote_Panel_DB_4".L2_OK AND "Remote_Panel_DB_5".L2_OK AND NOT "L3_Estop" AND NOT "Shuttle_EStop_All" AND "Lock_8_Estop_CH1" AND "Lock_11_Estop_CH1";
   "L4_OK" := "Remote_Panel_DB_1".L4_OK AND "Remote_Panel_DB_2".L4_OK AND "Remote_Panel_DB_3".L4_OK AND "Remote_Panel_DB_4".L4_OK AND "Remote_Panel_DB_5".L4_OK AND "Main_Panel_DB".Main_Panel_OK AND "Remote_Panel_DB_1".L3_OK AND "Remote_Panel_DB_2".L3_OK AND "Remote_Panel_DB_3".L3_OK AND "Remote_Panel_DB_4".L3_OK AND "Remote_Panel_DB_5".L3_OK AND NOT "L4_Estop" AND NOT "Shuttle_EStop_All";
   "L5_OK" := "Remote_Panel_DB_1".L5_OK AND "Remote_Panel_DB_2".L5_OK AND "Remote_Panel_DB_3".L5_OK AND "Remote_Panel_DB_4".L5_OK AND "Remote_Panel_DB_5".L5_OK AND "Main_Panel_DB".Main_Panel_OK AND "Remote_Panel_DB_1".L4_OK AND "Remote_Panel_DB_2".L4_OK AND "Remote_Panel_DB_3".L4_OK AND "Remote_Panel_DB_4".L4_OK AND "Remote_Panel_DB_5".L4_OK AND NOT "L5_Estop" AND NOT "Shuttle_EStop_All";
   "L6_OK" := "Remote_Panel_DB_1".L6_OK AND "Remote_Panel_DB_2".L6_OK AND "Remote_Panel_DB_3".L6_OK AND "Remote_Panel_DB_4".L6_OK AND "Remote_Panel_DB_5".L6_OK AND "Main_Panel_DB".Main_Panel_OK AND "Remote_Panel_DB_1".L5_OK AND "Remote_Panel_DB_2".L5_OK AND "Remote_Panel_DB_3".L5_OK AND "Remote_Panel_DB_4".L5_OK AND "Remote_Panel_DB_5".L4_OK AND NOT "L6_Estop" AND NOT "Shuttle_EStop_All";
   "L7_OK" := "Remote_Panel_DB_1".L7_OK AND "Remote_Panel_DB_2".L7_OK AND "Remote_Panel_DB_3".L7_OK AND "Remote_Panel_DB_4".L7_OK AND "Remote_Panel_DB_5".L7_OK AND "Main_Panel_DB".Main_Panel_OK AND "Remote_Panel_DB_1".L6_OK AND "Remote_Panel_DB_2".L6_OK AND "Remote_Panel_DB_3".L6_OK AND "Remote_Panel_DB_4".L6_OK AND "Remote_Panel_DB_5".L6_OK AND NOT "L7_Estop" AND NOT "Shuttle_EStop_All";
   "L8_OK" := "Remote_Panel_DB_1".L8_OK AND "Remote_Panel_DB_2".L8_OK AND "Remote_Panel_DB_3".L8_OK AND "Remote_Panel_DB_4".L8_OK AND "Remote_Panel_DB_5".L8_OK AND "Main_Panel_DB".Main_Panel_OK AND "Remote_Panel_DB_1".L7_OK AND "Remote_Panel_DB_2".L7_OK AND "Remote_Panel_DB_3".L7_OK AND "Remote_Panel_DB_4".L7_OK AND "Remote_Panel_DB_5".L7_OK AND NOT "L8_Estop" AND NOT "Shuttle_EStop_All";
END_REGION

REGION Network 10: LOCKS
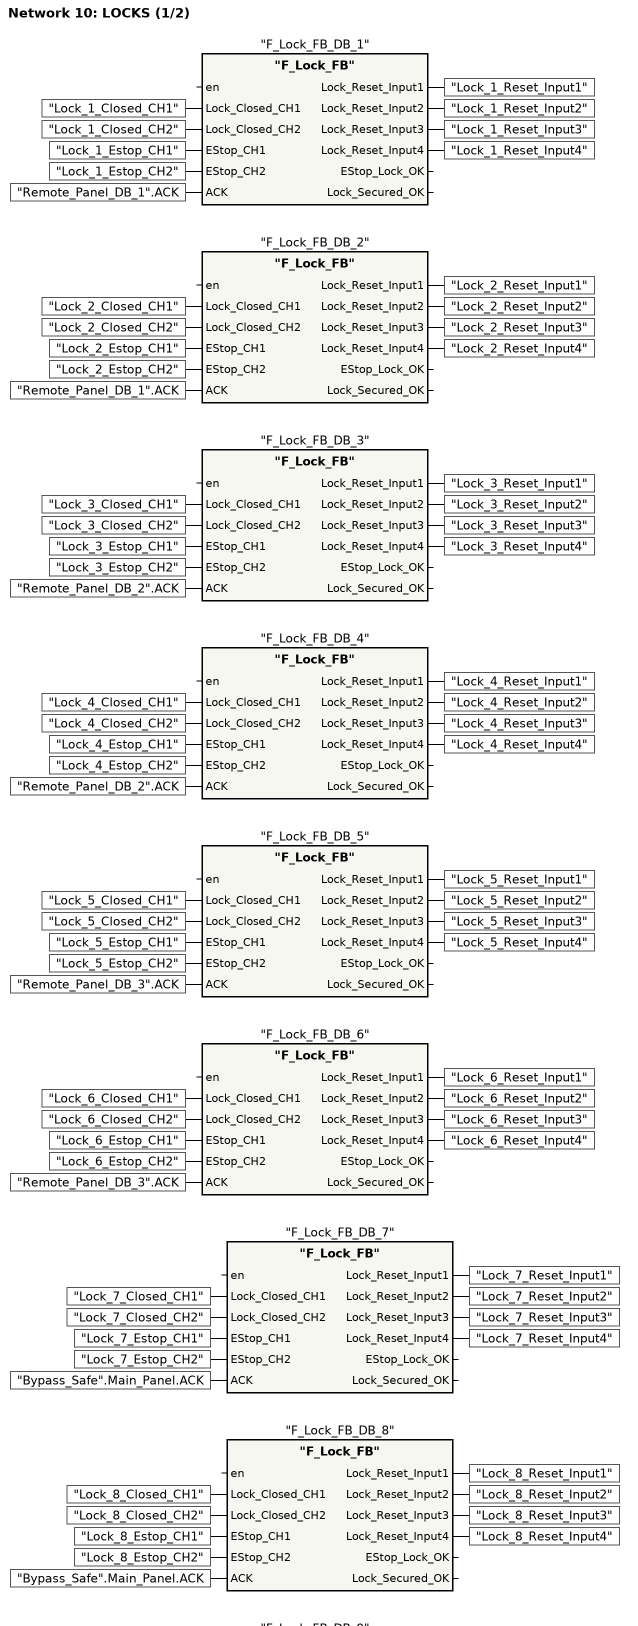
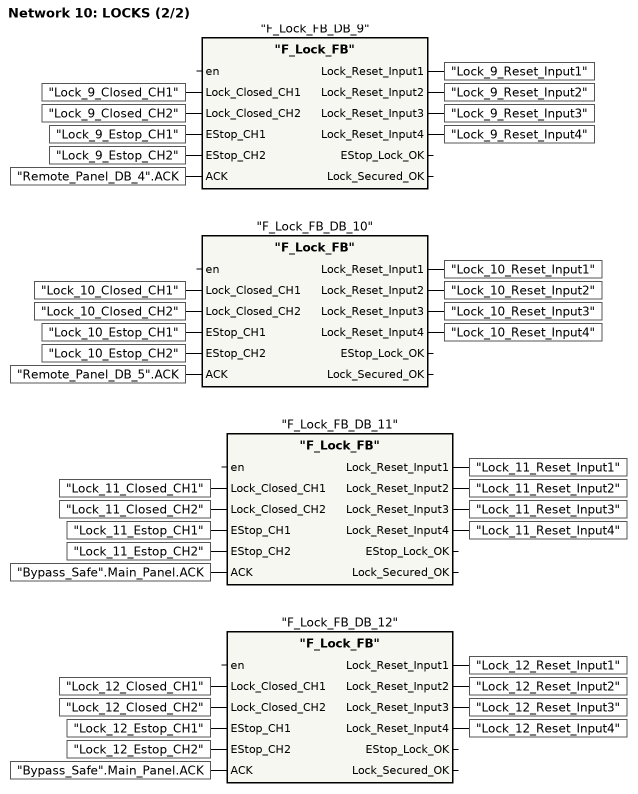
   "F_Lock_FB_DB_1"(Lock_Closed_CH1 := "Lock_1_Closed_CH1",   // "F_Lock_FB"
                    Lock_Closed_CH2 := "Lock_1_Closed_CH2",
                    EStop_CH1 := "Lock_1_Estop_CH1",
                    EStop_CH2 := "Lock_1_Estop_CH2",
                    ACK := "Remote_Panel_DB_1".ACK,
                    Lock_Reset_Input1 => "Lock_1_Reset_Input1",
                    Lock_Reset_Input2 => "Lock_1_Reset_Input2",
                    Lock_Reset_Input3 => "Lock_1_Reset_Input3",
                    Lock_Reset_Input4 => "Lock_1_Reset_Input4");
   "F_Lock_FB_DB_2"(Lock_Closed_CH1 := "Lock_2_Closed_CH1",   // "F_Lock_FB"
                    Lock_Closed_CH2 := "Lock_2_Closed_CH2",
                    EStop_CH1 := "Lock_2_Estop_CH1",
                    EStop_CH2 := "Lock_2_Estop_CH2",
                    ACK := "Remote_Panel_DB_1".ACK,
                    Lock_Reset_Input1 => "Lock_2_Reset_Input1",
                    Lock_Reset_Input2 => "Lock_2_Reset_Input2",
                    Lock_Reset_Input3 => "Lock_2_Reset_Input3",
                    Lock_Reset_Input4 => "Lock_2_Reset_Input4");
   "F_Lock_FB_DB_3"(Lock_Closed_CH1 := "Lock_3_Closed_CH1",   // "F_Lock_FB"
                    Lock_Closed_CH2 := "Lock_3_Closed_CH2",
                    EStop_CH1 := "Lock_3_Estop_CH1",
                    EStop_CH2 := "Lock_3_Estop_CH2",
                    ACK := "Remote_Panel_DB_2".ACK,
                    Lock_Reset_Input1 => "Lock_3_Reset_Input1",
                    Lock_Reset_Input2 => "Lock_3_Reset_Input2",
                    Lock_Reset_Input3 => "Lock_3_Reset_Input3",
                    Lock_Reset_Input4 => "Lock_3_Reset_Input4");
   "F_Lock_FB_DB_4"(Lock_Closed_CH1 := "Lock_4_Closed_CH1",   // "F_Lock_FB"
                    Lock_Closed_CH2 := "Lock_4_Closed_CH2",
                    EStop_CH1 := "Lock_4_Estop_CH1",
                    EStop_CH2 := "Lock_4_Estop_CH2",
                    ACK := "Remote_Panel_DB_2".ACK,
                    Lock_Reset_Input1 => "Lock_4_Reset_Input1",
                    Lock_Reset_Input2 => "Lock_4_Reset_Input2",
                    Lock_Reset_Input3 => "Lock_4_Reset_Input3",
                    Lock_Reset_Input4 => "Lock_4_Reset_Input4");
   "F_Lock_FB_DB_5"(Lock_Closed_CH1 := "Lock_5_Closed_CH1",   // "F_Lock_FB"
                    Lock_Closed_CH2 := "Lock_5_Closed_CH2",
                    EStop_CH1 := "Lock_5_Estop_CH1",
                    EStop_CH2 := "Lock_5_Estop_CH2",
                    ACK := "Remote_Panel_DB_3".ACK,
                    Lock_Reset_Input1 => "Lock_5_Reset_Input1",
                    Lock_Reset_Input2 => "Lock_5_Reset_Input2",
                    Lock_Reset_Input3 => "Lock_5_Reset_Input3",
                    Lock_Reset_Input4 => "Lock_5_Reset_Input4");
   "F_Lock_FB_DB_6"(Lock_Closed_CH1 := "Lock_6_Closed_CH1",   // "F_Lock_FB"
                    Lock_Closed_CH2 := "Lock_6_Closed_CH2",
                    EStop_CH1 := "Lock_6_Estop_CH1",
                    EStop_CH2 := "Lock_6_Estop_CH2",
                    ACK := "Remote_Panel_DB_3".ACK,
                    Lock_Reset_Input1 => "Lock_6_Reset_Input1",
                    Lock_Reset_Input2 => "Lock_6_Reset_Input2",
                    Lock_Reset_Input3 => "Lock_6_Reset_Input3",
                    Lock_Reset_Input4 => "Lock_6_Reset_Input4");
   "F_Lock_FB_DB_7"(Lock_Closed_CH1 := "Lock_7_Closed_CH1",   // "F_Lock_FB"
                    Lock_Closed_CH2 := "Lock_7_Closed_CH2",
                    EStop_CH1 := "Lock_7_Estop_CH1",
                    EStop_CH2 := "Lock_7_Estop_CH2",
                    ACK := "Bypass_Safe".Main_Panel.ACK,
                    Lock_Reset_Input1 => "Lock_7_Reset_Input1",
                    Lock_Reset_Input2 => "Lock_7_Reset_Input2",
                    Lock_Reset_Input3 => "Lock_7_Reset_Input3",
                    Lock_Reset_Input4 => "Lock_7_Reset_Input4");
   "F_Lock_FB_DB_8"(Lock_Closed_CH1 := "Lock_8_Closed_CH1",   // "F_Lock_FB"
                    Lock_Closed_CH2 := "Lock_8_Closed_CH2",
                    EStop_CH1 := "Lock_8_Estop_CH1",
                    EStop_CH2 := "Lock_8_Estop_CH2",
                    ACK := "Bypass_Safe".Main_Panel.ACK,
                    Lock_Reset_Input1 => "Lock_8_Reset_Input1",
                    Lock_Reset_Input2 => "Lock_8_Reset_Input2",
                    Lock_Reset_Input3 => "Lock_8_Reset_Input3",
                    Lock_Reset_Input4 => "Lock_8_Reset_Input4");
   "F_Lock_FB_DB_9"(Lock_Closed_CH1 := "Lock_9_Closed_CH1",   // "F_Lock_FB"
                    Lock_Closed_CH2 := "Lock_9_Closed_CH2",
                    EStop_CH1 := "Lock_9_Estop_CH1",
                    EStop_CH2 := "Lock_9_Estop_CH2",
                    ACK := "Remote_Panel_DB_4".ACK,
                    Lock_Reset_Input1 => "Lock_9_Reset_Input1",
                    Lock_Reset_Input2 => "Lock_9_Reset_Input2",
                    Lock_Reset_Input3 => "Lock_9_Reset_Input3",
                    Lock_Reset_Input4 => "Lock_9_Reset_Input4");
   "F_Lock_FB_DB_10"(Lock_Closed_CH1 := "Lock_10_Closed_CH1",   // "F_Lock_FB"
                     Lock_Closed_CH2 := "Lock_10_Closed_CH2",
                     EStop_CH1 := "Lock_10_Estop_CH1",
                     EStop_CH2 := "Lock_10_Estop_CH2",
                     ACK := "Remote_Panel_DB_5".ACK,
                     Lock_Reset_Input1 => "Lock_10_Reset_Input1",
                     Lock_Reset_Input2 => "Lock_10_Reset_Input2",
                     Lock_Reset_Input3 => "Lock_10_Reset_Input3",
                     Lock_Reset_Input4 => "Lock_10_Reset_Input4");
   "F_Lock_FB_DB_11"(Lock_Closed_CH1 := "Lock_11_Closed_CH1",   // "F_Lock_FB"
                     Lock_Closed_CH2 := "Lock_11_Closed_CH2",
                     EStop_CH1 := "Lock_11_Estop_CH1",
                     EStop_CH2 := "Lock_11_Estop_CH2",
                     ACK := "Bypass_Safe".Main_Panel.ACK,
                     Lock_Reset_Input1 => "Lock_11_Reset_Input1",
                     Lock_Reset_Input2 => "Lock_11_Reset_Input2",
                     Lock_Reset_Input3 => "Lock_11_Reset_Input3",
                     Lock_Reset_Input4 => "Lock_11_Reset_Input4");
   "F_Lock_FB_DB_12"(Lock_Closed_CH1 := "Lock_12_Closed_CH1",   // "F_Lock_FB"
                     Lock_Closed_CH2 := "Lock_12_Closed_CH2",
                     EStop_CH1 := "Lock_12_Estop_CH1",
                     EStop_CH2 := "Lock_12_Estop_CH2",
                     ACK := "Bypass_Safe".Main_Panel.ACK,
                     Lock_Reset_Input1 => "Lock_12_Reset_Input1",
                     Lock_Reset_Input2 => "Lock_12_Reset_Input2",
                     Lock_Reset_Input3 => "Lock_12_Reset_Input3",
                     Lock_Reset_Input4 => "Lock_12_Reset_Input4");
END_REGION

REGION Network 11: Safety OK
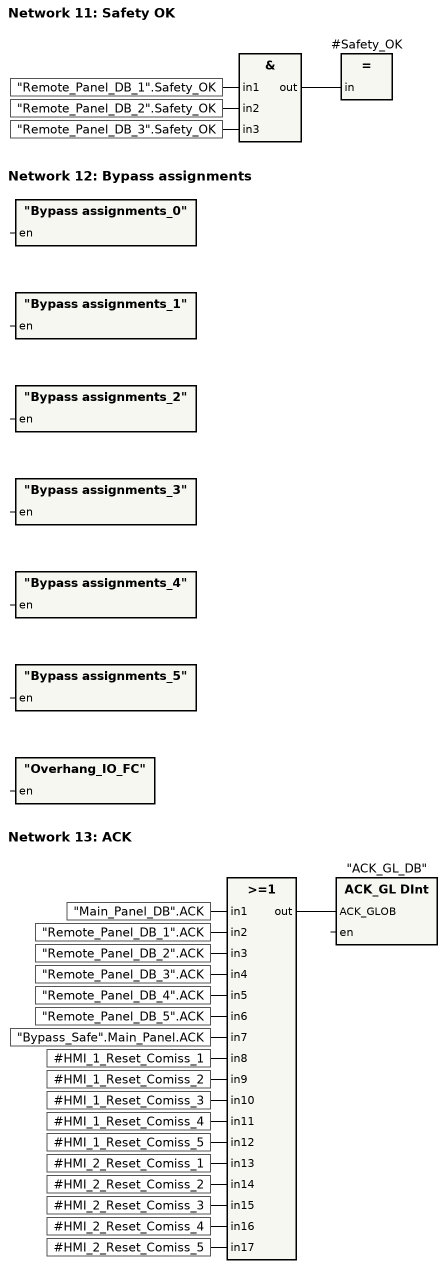
   #Safety_OK := "Remote_Panel_DB_1".Safety_OK AND "Remote_Panel_DB_2".Safety_OK AND "Remote_Panel_DB_3".Safety_OK;
END_REGION

REGION Network 12: Bypass assignments
   "Bypass assignments_0"();
   "Bypass assignments_1"();
   "Bypass assignments_2"();
   "Bypass assignments_3"();
   "Bypass assignments_4"();
   "Bypass assignments_5"();
   "Overhang_IO_FC"();
END_REGION

REGION Network 13: ACK
   "ACK_GL_DB"(ACK_GLOB := "Main_Panel_DB".ACK OR "Remote_Panel_DB_1".ACK OR "Remote_Panel_DB_2".ACK OR "Remote_Panel_DB_3".ACK OR "Remote_Panel_DB_4".ACK OR "Remote_Panel_DB_5".ACK OR "Bypass_Safe".Main_Panel.ACK OR #HMI_1_Reset_Comiss_1 OR #HMI_1_Reset_Comiss_2 OR #HMI_1_Reset_Comiss_3 OR #HMI_1_Reset_Comiss_4 OR #HMI_1_Reset_Comiss_5 OR #HMI_2_Reset_Comiss_1 OR #HMI_2_Reset_Comiss_2 OR #HMI_2_Reset_Comiss_3 OR #HMI_2_Reset_Comiss_4 OR #HMI_2_Reset_Comiss_5);   // ACK_GL
END_REGION

REGION Network 14: RESET PLC HMI
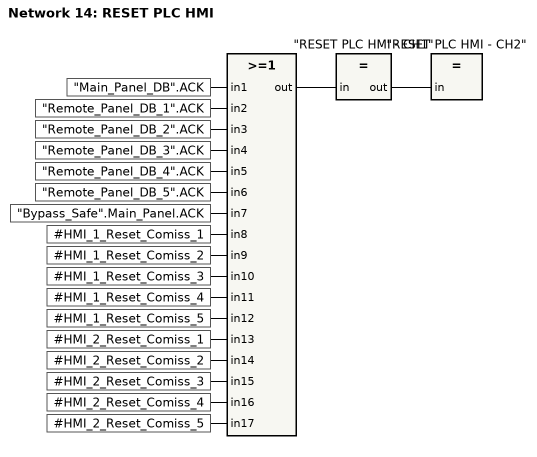
   "RESET PLC HMI - CH1" := "Main_Panel_DB".ACK OR "Remote_Panel_DB_1".ACK OR "Remote_Panel_DB_2".ACK OR "Remote_Panel_DB_3".ACK OR "Remote_Panel_DB_4".ACK OR "Remote_Panel_DB_5".ACK OR "Bypass_Safe".Main_Panel.ACK OR #HMI_1_Reset_Comiss_1 OR #HMI_1_Reset_Comiss_2 OR #HMI_1_Reset_Comiss_3 OR #HMI_1_Reset_Comiss_4 OR #HMI_1_Reset_Comiss_5 OR #HMI_2_Reset_Comiss_1 OR #HMI_2_Reset_Comiss_2 OR #HMI_2_Reset_Comiss_3 OR #HMI_2_Reset_Comiss_4 OR #HMI_2_Reset_Comiss_5;
   "RESET PLC HMI - CH2" := "RESET PLC HMI - CH1";
END_REGION
END_FUNCTION_BLOCK

FUNCTION_BLOCK "Remote_Panel"   // FB17, F_LAD
{ S7_Optimized_Access := 'TRUE' }
VERSION : 0.1
// stored: AutoNumber true, IsIECCheckEnabled false, UDAEnableTagReadback false
   VAR_INPUT
      ID : Int;
      Overtravel_Lower_limit : Bool;
      Overtravel_Upper_limit : Bool;
      Estop : Bool;
      Reset : Bool;
      Chain_Slack_1 : Bool;
      Chain_Slack_2 : Bool;
      Chain_Slack_3 : Bool;
      Chain_Slack_4 : Bool;
      "Light Guards CX101" : Bool;
      "Light Guards CX201" : Bool;
      Gate_1 : Bool;
      Gate_2 : Bool;
      EStop_Lock_1 : Bool;
      EStop_Lock_2 : Bool;
      Lock_Secured_1 : Bool;
      Lock_Secured_2 : Bool;
      "EStop Level 1" : Bool;
      "EStop Level 2" : Bool;
      "EStop Level 3" : Bool;
      "EStop Level 4" : Bool;
      "EStop Level 5" : Bool;
      "EStop Level 6" : Bool;
      "EStop Level 7" : Bool;
      "EStop Level 8" : Bool;
      Bypass : "F_Bypass_RemotePanel";
      Material_Selection_1 : Bool;
      MR_1 : Bool;
      Material_Selection_2 : Bool;
      MR_2 : Bool;
      Overhang_Left : Bool;
      Overhang_Right : Bool;
   END_VAR
   VAR_OUTPUT
      Safety_OK : Bool;
      Bypass_Warning : Bool;
      "STO VTD - CH1" : Bool;
      "STO VTD - CH2" : Bool;
      "STO CONVEYOR VTD - CH1" : Bool;
      "STO CONVEYOR VTD - CH2" : Bool;
      "STO CNV VFD (Level 1,2,3 - Side1) - CH1" : Bool;
      "STO CNV VFD (Level 1,2,3 - Side1) - CH2" : Bool;
      "STO CNV VFD (Level 1,2,3 - Side2) - CH1" : Bool;
      "STO CNV VFD (Level 1,2,3 - Side2) - CH2" : Bool;
      "STO CNV VFD (Level 4,5,6 - Side1) - CH1" : Bool;
      "STO CNV VFD (Level 4,5,6 - Side1) - CH2" : Bool;
      "STO CNV VFD (Level 4,5,6 - Side2) - CH1" : Bool;
      "STO CNV VFD (Level 4,5,6 - Side2) - CH2" : Bool;
      "STO CNV VFD (Level 7,8 - Side1) - CH1" : Bool;
      "STO CNV VFD (Level 7,8 - Side1) - CH2" : Bool;
      "STO CNV VFD (Level 7,8 - Side2) - CH1" : Bool;
      "STO CNV VFD (Level 7,8 - Side2) - CH2" : Bool;
      "Power Enable Safety Stopper Conveyors (Level 1,2,3 - Side1) - CH1" : Bool;
      "Power Enable Safety Stopper Conveyors (Level 1,2,3 - Side1) - CH2" : Bool;
      "Power Enable Safety Stopper Conveyors (Level 1,2,3 - Side2) - CH1" : Bool;
      "Power Enable Safety Stopper Conveyors (Level 1,2,3 - Side2) - CH2" : Bool;
      "Power Enable Safety Stopper Conveyors (Level 4,5,6 - Side1) - CH1" : Bool;
      "Power Enable Safety Stopper Conveyors (Level 4,5,6 - Side1) - CH2" : Bool;
      "Power Enable Safety Stopper Conveyors (Level 4,5,6 - Side2) - CH1" : Bool;
      "Power Enable Safety Stopper Conveyors (Level 4,5,6 - Side2) - CH2" : Bool;
      "Power Enable Safety Stopper Conveyors (Level 7,8 - Side1) - CH1" : Bool;
      "Power Enable Safety Stopper Conveyors (Level 7,8 - Side1) - CH2" : Bool;
      "Power Enable Safety Stopper Conveyors (Level 7,8 - Side2) - CH1" : Bool;
      "Power Enable Safety Stopper Conveyors (Level 7,8 - Side2) - CH2" : Bool;
      "VTU Hoist Brake Sfty Enable - CH1" : Bool;
      "VTU Hoist Brake Sfty Enable - CH2" : Bool;
      ACK { ExternalAccessible := 'False'; ExternalVisible := 'False'; ExternalWritable := 'False'} : Bool;
      L1_OK : Bool;
      L2_OK : Bool;
      L3_OK : Bool;
      L4_OK : Bool;
      L5_OK : Bool;
      L6_OK : Bool;
      L7_OK : Bool;
      L8_OK : Bool;
      EStop_Lock_1_OK : Bool;
      EStop_Lock_2_OK : Bool;
      Lock_Secured_1_OK : Bool;
      Lock_Secured_2_OK : Bool;
      Safety_Ok_Conf : Bool;
   END_VAR
   VAR
      Overtravel_Lower_Limit_DB : ESTOP1;
      Overtravel_Upper_Limit_DB : ESTOP1;
      Estop_Cabinet_DB : ESTOP1;
      Chain_Slack_1_DB : ESTOP1;
      Chain_Slack_2_DB : ESTOP1;
      Chain_Slack_3_DB : ESTOP1;
      Chain_Slack_4_DB : ESTOP1;
      Light_Guards_CX101 : ESTOP1;
      Light_Guards_CX201 : ESTOP1;
      Gate_1_DB : ESTOP1;
      Gate_2_DB : ESTOP1;
      EStop_Lock_1_DB : ESTOP1;
      EStop_Lock_2_DB : ESTOP1;
      Lock_Secured_1_DB : ESTOP1;
      Lock_Secured_2_DB : ESTOP1;
      "EStop Level 1_DB" : ESTOP1;
      "EStop Level 2_DB" : ESTOP1;
      "EStop Level 3_DB" : ESTOP1;
      "EStop Level 4_DB" : ESTOP1;
      "EStop Level 5_DB" : ESTOP1;
      "EStop Level 6_DB" : ESTOP1;
      "EStop Level 7_DB" : ESTOP1;
      "EStop Level 8_DB" : ESTOP1;
      Mute_LG_1_DB : "SICK Safe Entry Exit HW PLC V02";
      Distance_Materia_To_LG : DInt;
      Mute_LG_2_DB : "SICK Safe Entry Exit HW PLC V02";
      F_T_Delay_Sae_OK : TOF;
      F_T_Delay_CL_4 : TOF;
      F_T_Delay_CL_3 : TOF;
      F_T_Delay_CL_2 : TOF;
      F_T_Delay_CL_1 : TOF;
      Chain_Slack_1_Filtered { ExternalAccessible := 'False'; ExternalVisible := 'False'; ExternalWritable := 'False'} : Bool;
      Chain_Slack_2_Filtered { ExternalAccessible := 'False'; ExternalVisible := 'False'; ExternalWritable := 'False'} : Bool;
      Chain_Slack_3_Filtered { ExternalAccessible := 'False'; ExternalVisible := 'False'; ExternalWritable := 'False'} : Bool;
      Chain_Slack_4_Filtered { ExternalAccessible := 'False'; ExternalVisible := 'False'; ExternalWritable := 'False'} : Bool;
      Light_Guard_Tuned : Bool;
      Light_Guard_Tuned_Euro : Bool;
      Light_Guard_Tuned_UK : Bool;
      Light_Guard_Tuned_UK_Infeed : Bool;
      Light_Guard_Tuned_Euro_Infeed : Bool;
      Light_Guard_Tuned_Infeed : Bool;
      F_Timer_Infeed_UK : TP;
      F_Timer_Infeed_E : TP;
      F_Timer_Outfeed_UK : TP;
      F_Timer_Outfeed_E : TP;
      Overhang_Left_DB : ESTOP1;
      Overhang_Right_DB : ESTOP1;
   END_VAR
   VAR_TEMP
      EStop_Levels_OK : Bool;
   END_VAR
   VAR_TEMP   // added for the SCL form of the ladder/FBD networks
      _w1 : Bool;
   END_VAR
BEGIN

REGION Network 1: RESET CABINET
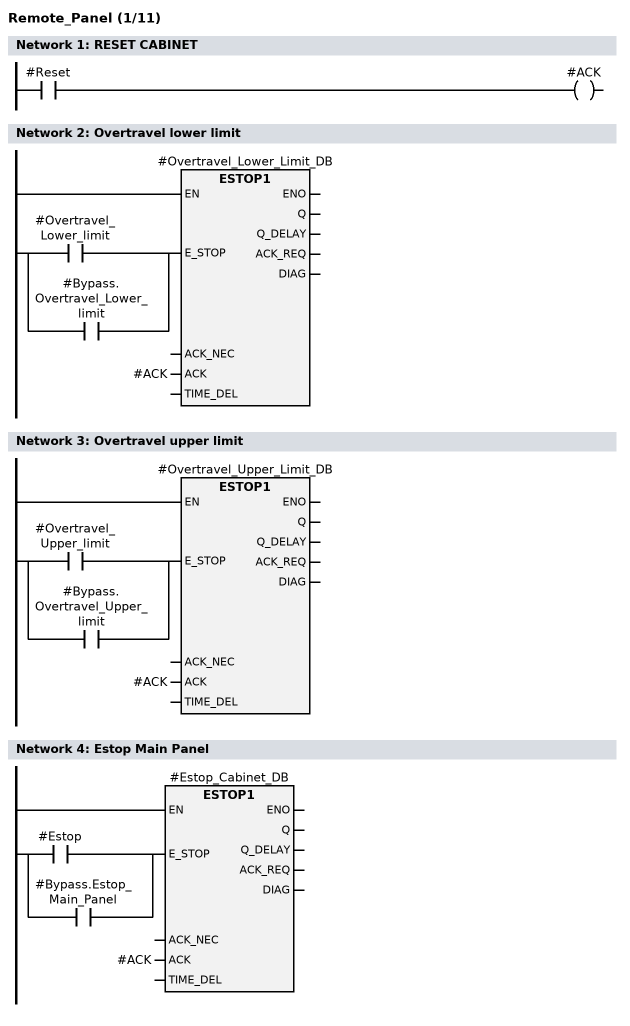
   RUNG wire#powerrail
      Contact( #Reset )
      Coil( #ACK )
   END_RUNG
   // the same network as SCL:
   #ACK := #Reset;
END_REGION

REGION Network 2: Overtravel lower limit
   RUNG wire#powerrail
      #Overtravel_Lower_Limit_DB.ESTOP1(E_STOP := wire#w1, ACK_NEC :=, ACK := #ACK, TIME_DEL :=, Q =>, Q_DELAY =>, ACK_REQ =>, DIAG =>)
   END_RUNG
   RUNG wire#powerrail
      Contact( #Overtravel_Lower_limit )
   END_RUNG wire#w1
   RUNG wire#powerrail
      Contact( #Bypass.Overtravel_Lower_limit )
   END_RUNG wire#w1
   // the same network as SCL:
   #Overtravel_Lower_Limit_DB(E_STOP := #Overtravel_Lower_limit OR #Bypass.Overtravel_Lower_limit, ACK := #ACK);   // ESTOP1
END_REGION

REGION Network 3: Overtravel upper limit
   RUNG wire#powerrail
      #Overtravel_Upper_Limit_DB.ESTOP1(E_STOP := wire#w1, ACK_NEC :=, ACK := #ACK, TIME_DEL :=, Q =>, Q_DELAY =>, ACK_REQ =>, DIAG =>)
   END_RUNG
   RUNG wire#powerrail
      Contact( #Overtravel_Upper_limit )
   END_RUNG wire#w1
   RUNG wire#powerrail
      Contact( #Bypass.Overtravel_Upper_limit )
   END_RUNG wire#w1
   // the same network as SCL:
   #Overtravel_Upper_Limit_DB(E_STOP := #Overtravel_Upper_limit OR #Bypass.Overtravel_Upper_limit, ACK := #ACK);   // ESTOP1
END_REGION

REGION Network 4: Estop Main Panel
   RUNG wire#powerrail
      #Estop_Cabinet_DB.ESTOP1(E_STOP := wire#w1, ACK_NEC :=, ACK := #ACK, TIME_DEL :=, Q =>, Q_DELAY =>, ACK_REQ =>, DIAG =>)
   END_RUNG
   RUNG wire#powerrail
      Contact( #Estop )
   END_RUNG wire#w1
   RUNG wire#powerrail
      Contact( #Bypass.Estop_Main_Panel )
   END_RUNG wire#w1
   // the same network as SCL:
   #Estop_Cabinet_DB(E_STOP := #Estop OR #Bypass.Estop_Main_Panel, ACK := #ACK);   // ESTOP1
END_REGION

REGION Network 5: Chain slack 1
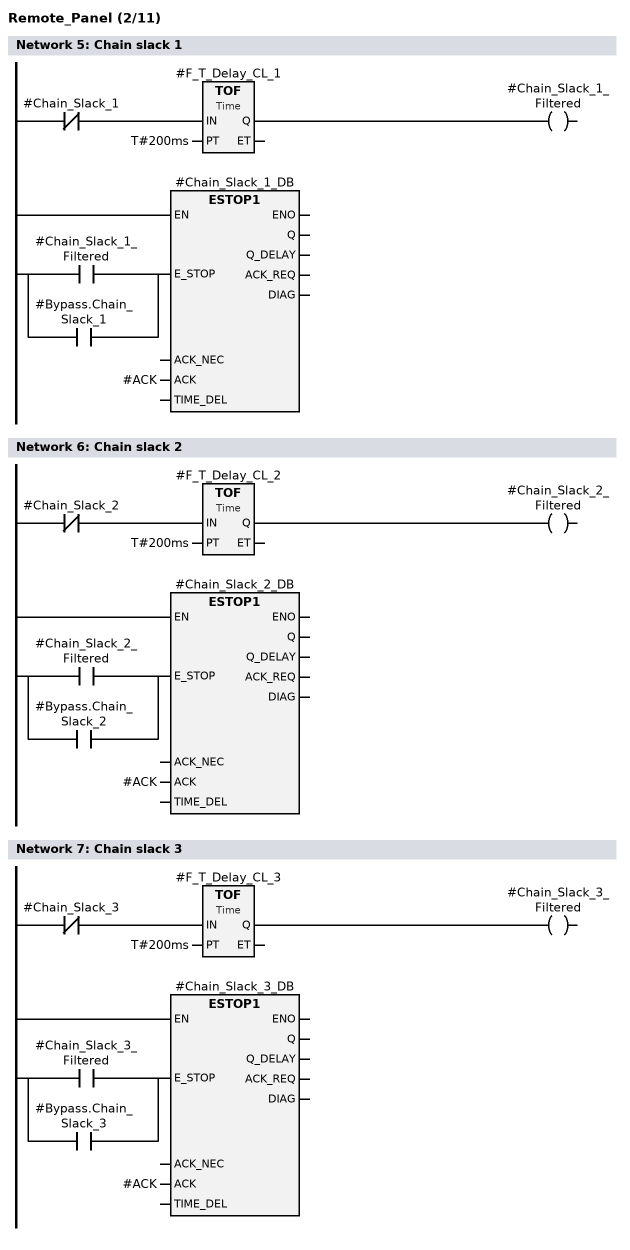
   RUNG wire#powerrail
      I_Contact( #Chain_Slack_1 )
      { S7_Templates := "[time_type := Time, codedbool_type := DInt]" } #F_T_Delay_CL_1.TOF(pt := T#200ms, et =>)
      Coil( #Chain_Slack_1_Filtered )
   END_RUNG
   RUNG wire#powerrail
      #Chain_Slack_1_DB.ESTOP1(E_STOP := wire#w1, ACK_NEC :=, ACK := #ACK, TIME_DEL :=, Q =>, Q_DELAY =>, ACK_REQ =>, DIAG =>)
   END_RUNG
   RUNG wire#powerrail
      Contact( #Chain_Slack_1_Filtered )
   END_RUNG wire#w1
   RUNG wire#powerrail
      Contact( #Bypass.Chain_Slack_1 )
   END_RUNG wire#w1
   // the same network as SCL:
   #F_T_Delay_CL_1.TOF(IN := NOT #Chain_Slack_1, PT := T#200ms);
   #Chain_Slack_1_Filtered := #F_T_Delay_CL_1.Q;
   #Chain_Slack_1_DB(E_STOP := #Chain_Slack_1_Filtered OR #Bypass.Chain_Slack_1, ACK := #ACK);   // ESTOP1
END_REGION

REGION Network 6: Chain slack 2
   RUNG wire#powerrail
      I_Contact( #Chain_Slack_2 )
      { S7_Templates := "[time_type := Time, codedbool_type := DInt]" } #F_T_Delay_CL_2.TOF(pt := T#200ms, et =>)
      Coil( #Chain_Slack_2_Filtered )
   END_RUNG
   RUNG wire#powerrail
      #Chain_Slack_2_DB.ESTOP1(E_STOP := wire#w1, ACK_NEC :=, ACK := #ACK, TIME_DEL :=, Q =>, Q_DELAY =>, ACK_REQ =>, DIAG =>)
   END_RUNG
   RUNG wire#powerrail
      Contact( #Chain_Slack_2_Filtered )
   END_RUNG wire#w1
   RUNG wire#powerrail
      Contact( #Bypass.Chain_Slack_2 )
   END_RUNG wire#w1
   // the same network as SCL:
   #F_T_Delay_CL_2.TOF(IN := NOT #Chain_Slack_2, PT := T#200ms);
   #Chain_Slack_2_Filtered := #F_T_Delay_CL_2.Q;
   #Chain_Slack_2_DB(E_STOP := #Chain_Slack_2_Filtered OR #Bypass.Chain_Slack_2, ACK := #ACK);   // ESTOP1
END_REGION

REGION Network 7: Chain slack 3
   RUNG wire#powerrail
      I_Contact( #Chain_Slack_3 )
      { S7_Templates := "[time_type := Time, codedbool_type := DInt]" } #F_T_Delay_CL_3.TOF(pt := T#200ms, et =>)
      Coil( #Chain_Slack_3_Filtered )
   END_RUNG
   RUNG wire#powerrail
      #Chain_Slack_3_DB.ESTOP1(E_STOP := wire#w1, ACK_NEC :=, ACK := #ACK, TIME_DEL :=, Q =>, Q_DELAY =>, ACK_REQ =>, DIAG =>)
   END_RUNG
   RUNG wire#powerrail
      Contact( #Chain_Slack_3_Filtered )
   END_RUNG wire#w1
   RUNG wire#powerrail
      Contact( #Bypass.Chain_Slack_3 )
   END_RUNG wire#w1
   // the same network as SCL:
   #F_T_Delay_CL_3.TOF(IN := NOT #Chain_Slack_3, PT := T#200ms);
   #Chain_Slack_3_Filtered := #F_T_Delay_CL_3.Q;
   #Chain_Slack_3_DB(E_STOP := #Chain_Slack_3_Filtered OR #Bypass.Chain_Slack_3, ACK := #ACK);   // ESTOP1
END_REGION

REGION Network 8: Chain slack 4
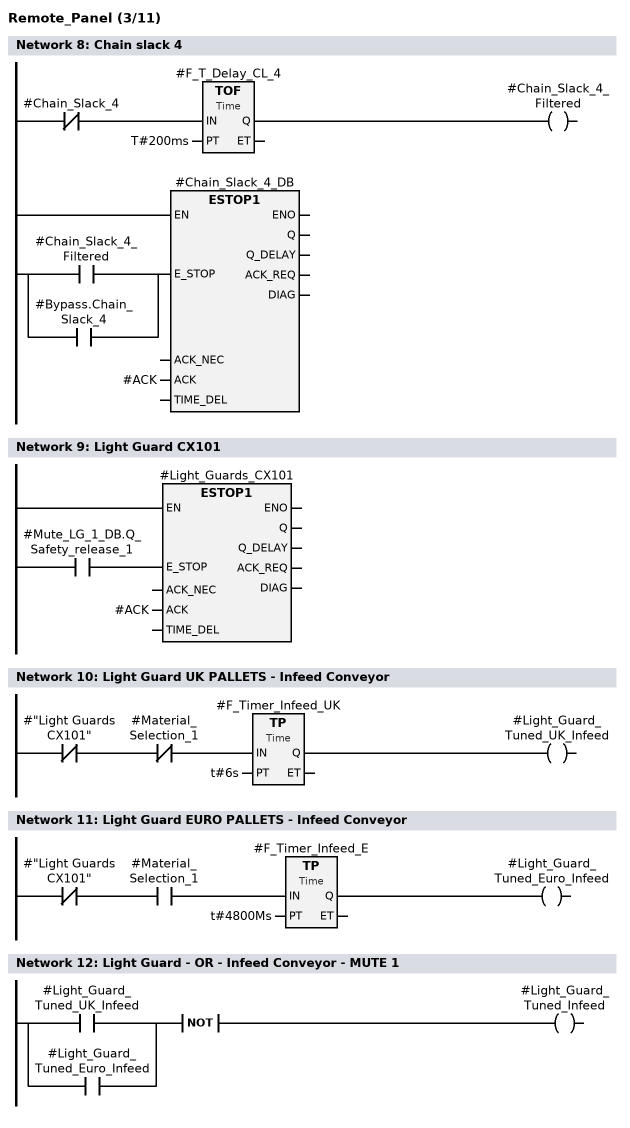
   RUNG wire#powerrail
      I_Contact( #Chain_Slack_4 )
      { S7_Templates := "[time_type := Time, codedbool_type := DInt]" } #F_T_Delay_CL_4.TOF(pt := T#200ms, et =>)
      Coil( #Chain_Slack_4_Filtered )
   END_RUNG
   RUNG wire#powerrail
      #Chain_Slack_4_DB.ESTOP1(E_STOP := wire#w1, ACK_NEC :=, ACK := #ACK, TIME_DEL :=, Q =>, Q_DELAY =>, ACK_REQ =>, DIAG =>)
   END_RUNG
   RUNG wire#powerrail
      Contact( #Chain_Slack_4_Filtered )
   END_RUNG wire#w1
   RUNG wire#powerrail
      Contact( #Bypass.Chain_Slack_4 )
   END_RUNG wire#w1
   // the same network as SCL:
   #F_T_Delay_CL_4.TOF(IN := NOT #Chain_Slack_4, PT := T#200ms);
   #Chain_Slack_4_Filtered := #F_T_Delay_CL_4.Q;
   #Chain_Slack_4_DB(E_STOP := #Chain_Slack_4_Filtered OR #Bypass.Chain_Slack_4, ACK := #ACK);   // ESTOP1
END_REGION

REGION Network 9: Light Guard CX101
   RUNG wire#powerrail
      #Light_Guards_CX101.ESTOP1(E_STOP := wire#w1, ACK_NEC :=, ACK := #ACK, TIME_DEL :=, Q =>, Q_DELAY =>, ACK_REQ =>, DIAG =>)
   END_RUNG
   RUNG wire#powerrail
      Contact( #Mute_LG_1_DB.Q_Safety_release_1 )
   END_RUNG wire#w1
   // the same network as SCL:
   #Light_Guards_CX101(E_STOP := #Mute_LG_1_DB.Q_Safety_release_1, ACK := #ACK);   // ESTOP1
END_REGION

REGION Network 10: Light Guard UK PALLETS - Infeed Conveyor
   RUNG wire#powerrail
      I_Contact( #"Light Guards CX101" )
      I_Contact( #Material_Selection_1 )
      { S7_Templates := "[time_type := Time, codedbool_type := DInt]" } #F_Timer_Infeed_UK.TP(pt := t#6s, et =>)
      Coil( #Light_Guard_Tuned_UK_Infeed )
   END_RUNG
   // the same network as SCL:
   #F_Timer_Infeed_UK.TP(IN := NOT #"Light Guards CX101" AND NOT #Material_Selection_1, PT := t#6s);
   #Light_Guard_Tuned_UK_Infeed := #F_Timer_Infeed_UK.Q;
END_REGION

REGION Network 11: Light Guard EURO PALLETS - Infeed Conveyor
   RUNG wire#powerrail
      I_Contact( #"Light Guards CX101" )
      Contact( #Material_Selection_1 )
      { S7_Templates := "[time_type := Time, codedbool_type := DInt]" } #F_Timer_Infeed_E.TP(pt := t#4800Ms, et =>)
      Coil( #Light_Guard_Tuned_Euro_Infeed )
   END_RUNG
   // the same network as SCL:
   #F_Timer_Infeed_E.TP(IN := NOT #"Light Guards CX101" AND #Material_Selection_1, PT := t#4800Ms);
   #Light_Guard_Tuned_Euro_Infeed := #F_Timer_Infeed_E.Q;
END_REGION

REGION Network 12: Light Guard - OR - Infeed Conveyor - MUTE 1
   RUNG wire#powerrail
      Contact( #Light_Guard_Tuned_UK_Infeed )
      wire#w1
      Not()
      Coil( #Light_Guard_Tuned_Infeed )
   END_RUNG
   RUNG wire#powerrail
      Contact( #Light_Guard_Tuned_Euro_Infeed )
   END_RUNG wire#w1
   // the same network as SCL:
   #Light_Guard_Tuned_Infeed := NOT (#Light_Guard_Tuned_UK_Infeed OR #Light_Guard_Tuned_Euro_Infeed);
END_REGION

REGION Network 13: MUTE 1
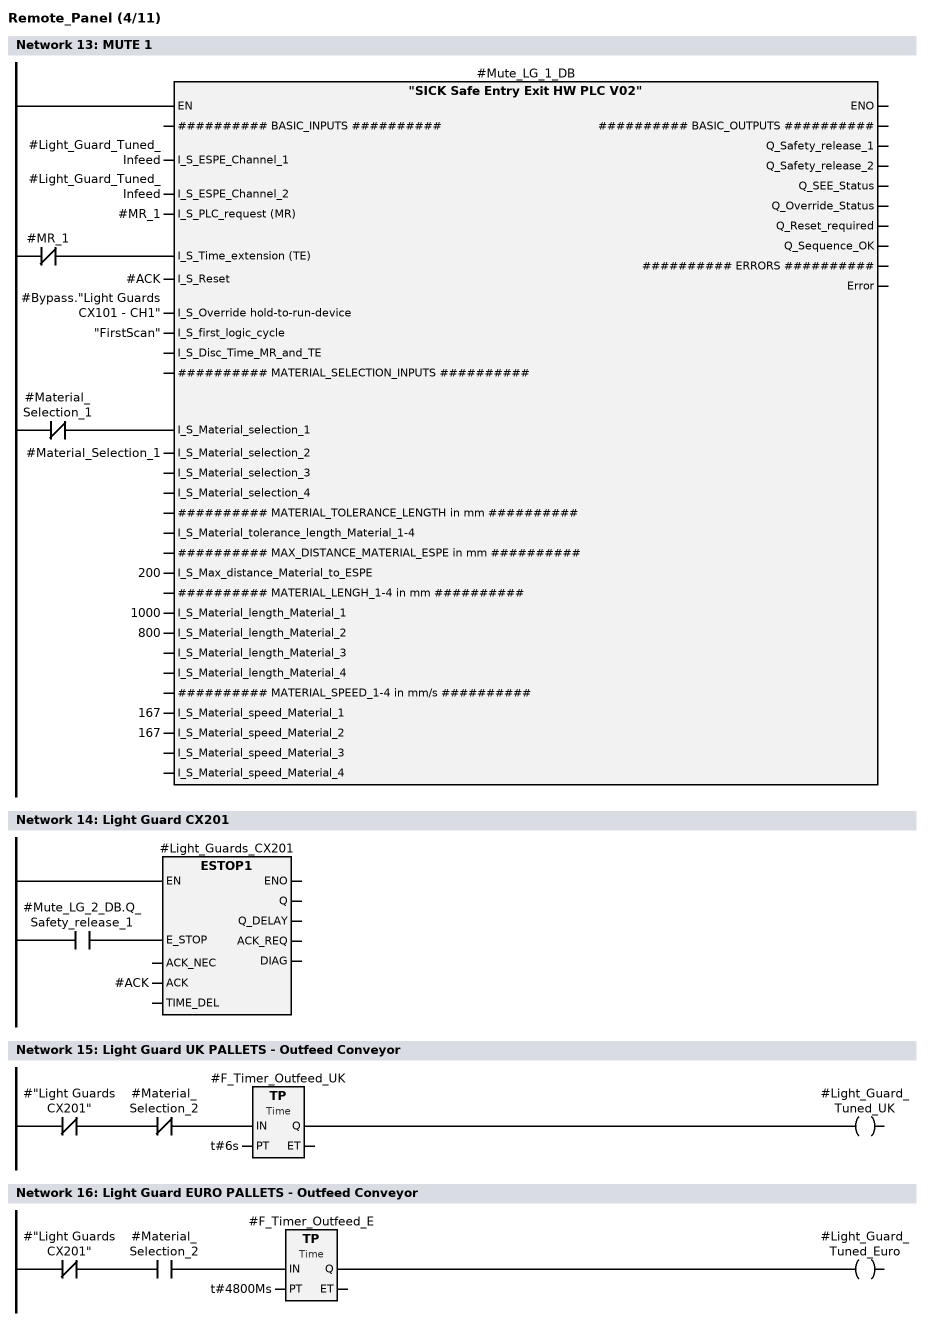
   RUNG wire#powerrail
      #Mute_LG_1_DB("I_S_Time_extension (TE)" := wire#w1, I_S_Material_selection_1 := wire#w2, "########## BASIC_INPUTS ##########" :=, I_S_ESPE_Channel_1 := #Light_Guard_Tuned_Infeed, I_S_ESPE_Channel_2 := #Light_Guard_Tuned_Infeed, "I_S_PLC_request (MR)" := #MR_1, I_S_Reset := #ACK, "I_S_Override hold-to-run-device" := #Bypass."Light Guards CX101 - CH1", I_S_first_logic_cycle := "FirstScan", I_S_Disc_Time_MR_and_TE :=, "########## MATERIAL_SELECTION_INPUTS ##########" :=, I_S_Material_selection_2 := #Material_Selection_1, I_S_Material_selection_3 :=, I_S_Material_selection_4 :=, "########## MATERIAL_TOLERANCE_LENGTH in mm ##########" :=, "I_S_Material_tolerance_length_Material_1-4" :=, "########## MAX_DISTANCE_MATERIAL_ESPE in mm ##########" :=, I_S_Max_distance_Material_to_ESPE := 200, "########## MATERIAL_LENGH_1-4 in mm ##########" :=, I_S_Material_length_Material_1 := 1000, I_S_Material_length_Material_2 := 800, I_S_Material_length_Material_3 :=, I_S_Material_length_Material_4 :=, "########## MATERIAL_SPEED_1-4 in mm/s ##########" :=, I_S_Material_speed_Material_1 := 167, I_S_Material_speed_Material_2 := 167, I_S_Material_speed_Material_3 :=, I_S_Material_speed_Material_4 :=, "########## BASIC_OUTPUTS ##########" =>, Q_Safety_release_1 =>, Q_Safety_release_2 =>, Q_SEE_Status =>, Q_Override_Status =>, Q_Reset_required =>, Q_Sequence_OK =>, "########## ERRORS ##########" =>, Error =>)
   END_RUNG
   RUNG wire#powerrail
      I_Contact( #MR_1 )
   END_RUNG wire#w1
   RUNG wire#powerrail
      I_Contact( #Material_Selection_1 )
   END_RUNG wire#w2
   // the same network as SCL:
   #Mute_LG_1_DB(I_S_ESPE_Channel_1 := #Light_Guard_Tuned_Infeed,   // "SICK Safe Entry Exit HW PLC V02"
                 I_S_ESPE_Channel_2 := #Light_Guard_Tuned_Infeed,
                 "I_S_PLC_request (MR)" := #MR_1,
                 "I_S_Time_extension (TE)" := NOT #MR_1,
                 I_S_Reset := #ACK,
                 "I_S_Override hold-to-run-device" := #Bypass."Light Guards CX101 - CH1",
                 I_S_first_logic_cycle := "FirstScan",
                 I_S_Material_selection_1 := NOT #Material_Selection_1,
                 I_S_Material_selection_2 := #Material_Selection_1,
                 I_S_Max_distance_Material_to_ESPE := 200,
                 I_S_Material_length_Material_1 := 1000,
                 I_S_Material_length_Material_2 := 800,
                 I_S_Material_speed_Material_1 := 167,
                 I_S_Material_speed_Material_2 := 167);
END_REGION

REGION Network 14: Light Guard CX201
   RUNG wire#powerrail
      #Light_Guards_CX201.ESTOP1(E_STOP := wire#w1, ACK_NEC :=, ACK := #ACK, TIME_DEL :=, Q =>, Q_DELAY =>, ACK_REQ =>, DIAG =>)
   END_RUNG
   RUNG wire#powerrail
      Contact( #Mute_LG_2_DB.Q_Safety_release_1 )
   END_RUNG wire#w1
   // the same network as SCL:
   #Light_Guards_CX201(E_STOP := #Mute_LG_2_DB.Q_Safety_release_1, ACK := #ACK);   // ESTOP1
END_REGION

REGION Network 15: Light Guard UK PALLETS - Outfeed Conveyor
   RUNG wire#powerrail
      I_Contact( #"Light Guards CX201" )
      I_Contact( #Material_Selection_2 )
      { S7_Templates := "[time_type := Time, codedbool_type := DInt]" } #F_Timer_Outfeed_UK.TP(pt := t#6s, et =>)
      Coil( #Light_Guard_Tuned_UK )
   END_RUNG
   // the same network as SCL:
   #F_Timer_Outfeed_UK.TP(IN := NOT #"Light Guards CX201" AND NOT #Material_Selection_2, PT := t#6s);
   #Light_Guard_Tuned_UK := #F_Timer_Outfeed_UK.Q;
END_REGION

REGION Network 16: Light Guard EURO PALLETS - Outfeed Conveyor
   RUNG wire#powerrail
      I_Contact( #"Light Guards CX201" )
      Contact( #Material_Selection_2 )
      { S7_Templates := "[time_type := Time, codedbool_type := DInt]" } #F_Timer_Outfeed_E.TP(pt := t#4800Ms, et =>)
      Coil( #Light_Guard_Tuned_Euro )
   END_RUNG
   // the same network as SCL:
   #F_Timer_Outfeed_E.TP(IN := NOT #"Light Guards CX201" AND #Material_Selection_2, PT := t#4800Ms);
   #Light_Guard_Tuned_Euro := #F_Timer_Outfeed_E.Q;
END_REGION

REGION Network 17: Light Guard - OR - Infeed Conveyor - MUTE 2
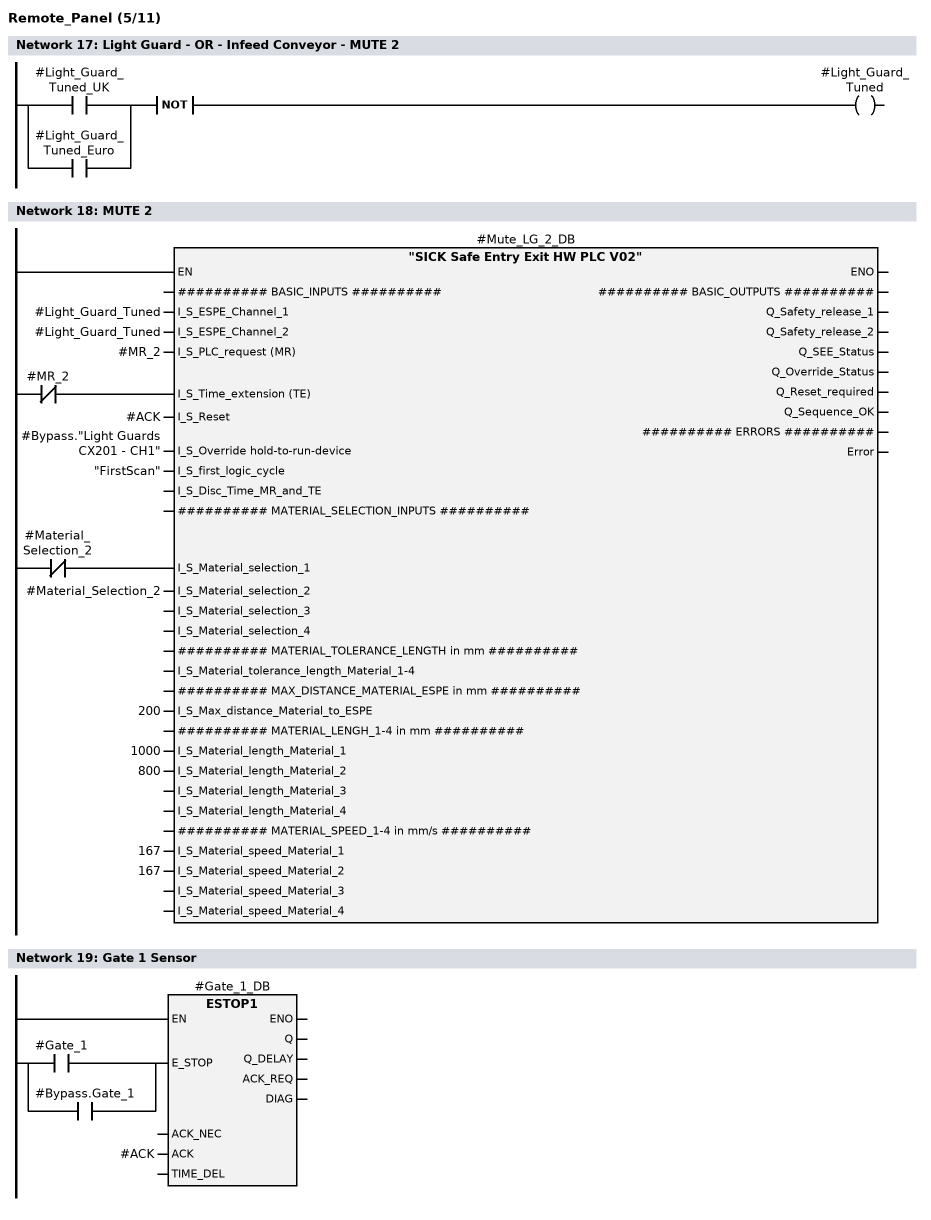
   RUNG wire#powerrail
      Contact( #Light_Guard_Tuned_UK )
      wire#w1
      Not()
      Coil( #Light_Guard_Tuned )
   END_RUNG
   RUNG wire#powerrail
      Contact( #Light_Guard_Tuned_Euro )
   END_RUNG wire#w1
   // the same network as SCL:
   #Light_Guard_Tuned := NOT (#Light_Guard_Tuned_UK OR #Light_Guard_Tuned_Euro);
END_REGION

